text list "EncoderแกนX (เบิกจ่าย)": 0 '0'; 1 '5935'; 2 '9155'; 3 '12375'; 4 '15595'; 5 '18815'; 6 '22035'; 7 '25255'; 8 '28475'; 9 '31695'; 10 '34915'; 11 '38135'; 12 '41355'; 13 '44575'; 14 '52483'; 15 '55703'; 16 '58923'; 17 '62143'; 18 '65363'; 19 '68583'; 20 '71803'; 21 '75023'; 22 '78243'; 23 '81463'; 24 '84683'; 25 '87903'; 26 '91123'; 27 '5935'; 28 '9155'; 29 '12375'; 30 '15595'; 31 '18815'; 32 '22035'; 33 '25255'; 34 '28475'; 35 '31695'; 36 '34915'; 37 '38135'; 38 '41355'; 39 '44575'; 40 '52483'; 41 '55703'; 42 '58923'; 43 '62143'; 44 '65363'; 45 '68583'; 46 '71803'; 47 '75023'; 48 '78243'; 49 '81463'; 50 '84683'; 51 '87903'; 52 '91123'; 53 '5935'; 54 '9155'; 55 '12375'; 56 '15595'; 57 '18815'; 58 '22035'; 59 '25255'; 60 '28475'; 61 '31695'; 62 '34915'; 63 '38135'; 64 '41355'; 65 '44575'; 66 '52483'; 67 '55703'; 68 '58923'; 69 '62143'; 70 '65363'; 71 '68583'; 72 '71803'; 73 '75023'; 74 '78243'; 75 '81463'; 76 '84683'; 77 '87903'; 78 '91123'; 79 '5935'; 80 '9155'; 81 '12375'; 82 '15595'; 83 '18815'; 84 '22035'; 85 '25255'; 86 '28475'; 87 '31695'; 88 '34915'; 89 '38135'; 90 '41355'; 91 '44575'; 92 '52483'; 93 '55703'; 94 '58923'; 95 '62143'; 96 '65363'; 97 '68583'; 98 '71803'; 99 '75023'; 100 '78243'; 101 '81463'; 102 '84683'; 103 '87903'; 104 '91123'; 105 '5935'; 106 '9155'; 107 '12375'; 108 '15595'; 109 '18815'; 110 '22035'; 111 '25255'; 112 '28475'; 113 '31695'; 114 '34915'; 115 '38135'; 116 '41355'; 117 '44575'; 118 '52483'; 119 '55703'; 120 '58923'; 121 '62143'; 122 '65363'; 123 '68583'; 124 '71803'; 125 '75023'; 126 '78243'; 127 '81463'; 128 '84683'; 129 '87903'; 130 '91123'; 131 '5935'; 132 '9155'; 133 '12375'; 134 '15595'; 135 '18815'; 136 '22035'; 137 '25255'; 138 '28475'; 139 '31695'; 140 '34915'; 141 '38135'; 142 '41355'; 143 '44575'; 144 '52483'; 145 '55703'; 146 '58923'; 147 '62143'; 148 '65363'; 149 '68583'; 150 '71803'; 151 '75023'; 152 '78243'; 153 '81463'; 154 '84683'; 155 '87903'; 156 '91123'; 157 '5935'; 158 '9155'; 159 '12375'; 160 '15595'; 161 '18815'; 162 '22035'; 163 '25255'; 164 '28475'; 165 '31695'; 166 '34915'; 167 '38135'; 168 '41355'; 169 '44575'; 170 '52483'; 171 '55703'; 172 '58923'; 173 '62143'; 174 '65363'; 175 '68583'; 176 '71803'; 177 '75023'; 178 '78243'; 179 '81463'; 180 '84683'; 181 '87903'; 182 '91123'; 183 '5935'; 184 '9155'; 185 '12375'; 186 '15595'; 187 '18815'; 188 '22035'; 189 '25255'; 190 '28475'; 191 '31695'; 192 '34915'; 193 '38135'; 194 '41355'; 195 '44575'; 196 '52483'; 197 '55703'; 198 '58923'; 199 '62143'; 200 '65363'; 201 '68583'; 202 '71803'; 203 '75023'; 204 '78243'; 205 '81463'; 206 '84683'; 207 '87903'; 208 '91123'; 209 '5935'; 210 '9155'; 211 '12375'; 212 '15595'; 213 '18815'; 214 '22035'; 215 '25255'; 216 '28475'; 217 '31695'; 218 '34915'; 219 '38135'; 220 '41355'; 221 '44575'; 222 '52483'; 223 '55703'; 224 '58923'; 225 '62143'; 226 '65363'; 227 '68583'; 228 '71803'; 229 '75023'; 230 '78243'; 231 '81463'; 232 '84683'; 233 '87903'; 234 '91123'; 235 '5935'; 236 '9155'; 237 '12375'; 238 '15595'; 239 '18815'; 240 '22035'; 241 '25255'; 242 '28475'; 243 '31695'; 244 '34915'; 245 '38135'; 246 '41355'; 247 '44575'; 248 '52483'; 249 '55703'; 250 '58923'; 251 '62143'; 252 '65363'; 253 '68583'; 254 '71803'; 255 '75023'; 256 '78243'; 257 '81463'; 258 '84683'; 259 '87903'; 260 '91123'; 261 '5935'; 262 '9155'; 263 '12375'; 264 '15595'; 265 '18815'; 266 '22035'; 267 '25255'; 268 '28475'; 269 '31695'; 270 '34915'; 271 '38135'; 272 '41355'; 273 '44575'; 274 '52483'; 275 '55703'; 276 '58923'; 277 '62143'; 278 '65363'; 279 '68583'; 280 '71803'; 281 '75023'; 282 '78243'; 283 '81463'; 284 '84683'; 285 '87903'; 286 '91123'; 287 '5935'; 288 '9155'; 289 '12375'; 290 '15595'; 291 '18815'; 292 '22035'; 293 '25255'; 294 '28475'; 295 '31695'; 296 '34915'; 297 '38135'; 298 '41355'; 299 '44575'; 300 '52483'; 301 '55703'; 302 '58923'; 303 '62143'; 304 '65363'; 305 '68583'; 306 '71803'; 307 '75023'; 308 '78243'; 309 '81463'; 310 '84683'; 311 '87903'; 312 '91123'; 313 '5935'; 314 '9155'; 315 '12375'; 316 '15595'; 317 '18815'; 318 '22035'; 319 '25255'; 320 '28475'; 321 '31695'; 322 '34915'; 323 '38135'; 324 '41355'; 325 '44575'; 326 '52483'; 327 '55703'; 328 '58923'; 329 '62143'; 330 '65363'; 331 '68583'; 332 '71803'; 333 '75023'; 334 '78243'; 335 '81463'; 336 '84683'; 337 '87903'; 338 '91123'; 339 '5935'; 340 '9155'; 341 '12375'; 342 '15595'; 343 '18815'; 344 '22035'; 345 '25255'; 346 '28475'; 347 '31695'; 348 '34915'; 349 '38135'; 350 '41355'; 351 '44575'; 352 '52483'; 353 '55703'; 354 '58923'; 355 '62143'; 356 '65363'; 357 '68583'; 358 '71803'; 359 '75023'; 360 '78243'; 361 '81463'; 362 '84683'; 363 '87903'; 364 '91123'; 365 '5935'; 366 '9155'; 367 '12375'; 368 '15595'; 369 '18815'; 370 '22035'; 371 '25255'; 372 '28475'; 373 '31695'; 374 '34915'; 375 '38135'; 376 '41355'; 377 '44575'; 378 '52483'; 379 '55703'; 380 '58923'; 381 '62143'; 382 '65363'; 383 '68583'; 384 '71803'; 385 '75023'; 386 '78243'; 387 '81463'; 388 '84683'; 389 '87903'; 390 '91123'; 391 '5935'; 392 '9155'; 393 '12375'; 394 '15595'; 395 '18815'; 396 '22035'; 397 '25255'; 398 '28475'; 399 '31695'; 400 '34915'; 401 '38135'; 402 '41355'; 403 '44575'; 404 '52483'; 405 '55703'; 406 '58923'; 407 '62143'; 408 '65363'; 409 '68583'; 410 '71803'; 411 '75023'; 412 '78243'; 413 '81463'; 414 '84683'; 415 '87903'; 416 '91123'; 417 '5935'; 418 '9155'; 419 '12375'; 420 '15595'; 421 '18815'; 422 '22035'; 423 '25255'; 424 '28475'; 425 '31695'; 426 '34915'; 427 '38135'; 428 '41355'; 429 '44575'; 430 '52483'; 431 '55703'; 432 '58923'; 433 '62143'; 434 '65363'; 435 '68583'; 436 '71803'; 437 '75023'; 438 '78243'; 439 '81463'; 440 '84683'; 441 '87903'; 442 '91123'; 443 '5935'; 444 '9155'; 445 '12375'; 446 '15595'; 447 '18815'; 448 '22035'; 449 '25255'; 450 '28475'; 451 '31695'; 452 '34915'; 453 '38135'; 454 '41355'; 455 '44575'; 456 '52483'; 457 '55703'; 458 '58923'; 459 '62143'; 460 '65363'; 461 '68583'; 462 '71803'; 463 '75023'; 464 '78243'; 465 '81463'; 466 '84683'; 467 '87903'; 468 '91123'; 469 '5935'; 470 '9155'; 471 '12375'; 472 '15595'; 473 '18815'; 474 '22035'; 475 '25255'; 476 '28475'; 477 '31695'; 478 '34915'; 479 '38135'; 480 '41355'; 481 '44575'; 482 '52483'; 483 '55703'; 484 '58923'; 485 '62143'; 486 '65363'; 487 '68583'; 488 '71803'; 489 '75023'; 490 '78243'; 491 '81463'; 492 '84683'; 493 '87903'; 494 '91123'

text list "Textlist_ScreenName": 1 'PROCESS OVERVIEW'; 5 'ALARMS'; 20 'ORDER'; 10 'SETTING'

text list "จัดเก็บ Motor speed1,2": 0 '0'; 1 '500'

text list "จัดเก็บ Current 1,2": 0 '0'; 1 '6'

text list "จัดเก็บ Power 1,2": 0 '0'; 1 '270'

text list "จัดเก็บVoltage 1,2": 0 '0'; 1 '66'

text list "จัดเก็บ Motor speed3": 0 '0'; 2 '1500'

text list "จัดเก็บ Current 3": 0 '0'; 2 '6'

text list "จัดเก็บ Power 3": 0 '0'; 2 '270'

text list "จัดเก็บVoltage 3": 0 '0'; 2 '66'

text list "เบิกจ่าย Motor speed1,2": 0 '0'; 1 '500'

text list "เบิกจ่าย Current 1,2": 0 '0'; 1 '6'

text list "เบิกจ่าย Power 1,2": 0 '0'; 1 '270'

text list "เบิกจ่ายVoltage 1,2": 0 '0'; 1 '66'

text list "เบิกจ่าย Motor speed3": 0 '0'; 2 '1500'

text list "เบิกจ่าย Current 3": 0 '0'; 2 '6'

text list "เบิกจ่าย Power 3": 0 '0'; 2 '270'

text list "เบิกจ่ายVoltage 3": 0 '0'; 2 '66'

text list "Status1": 0 'Stop'; 1 'Running'

graphic list "GriphList_Button_Start": 0 '-play-button-off'; 1 '-button-96-on'

graphic list "GriphList_Button_Setting": 0 'setting-green-off'; 1 'settings-96-off'

graphic list "GriphList_Button_Alarms": 0 'arning-96-off'; 1 'warning-96-on'

graphic list "GriphList_Button_Order": 0 'order-off'; 1 'order'

graphic list "GriphList_Button_Overview": 0 'overview-off'; 1 'overview-on'

PopupScreen "Confirm" 500x250
   TextField "Template_Text field_1" at 72,8 size 209x37; Text 'ยืนยันการสั่งซื้อ'
   Button "Button_1" at 426,9 size 64x32; TextOff 'X'
      on Click: function_efd93a16("Confirm", 0, 0, 0, -1, 1)
   GraphicView "Template_Graphic view_1" at 8,8 size 45x40; Picture "bell"
   GraphicView "Template_Graphic view_2" at 152,66 size 187x166; Picture "accept"

PopupScreen "ช่องยานี้เต็มแล้ว" 500x250
   TextField "Template_Text field_1" at 72,8 size 22x37; Text 'Text'
   Button "Button_1" at 426,9 size 64x32; TextOff 'X'
      on Click: function_efd93a16("ช่องยานี้เต็มแล้ว", 0, 0, 0, -1, 1)
   GraphicView "Template_Graphic view_1" at 8,8 size 45x40; Picture "bell"
   GraphicView "Template_Graphic view_2" at 152,66 size 187x166; Picture "close"

PopupScreen "จัดเก็บยาเสร็จสิ้น" 500x250
   TextField "Template_Text field_1" at 72,8 size 227x37; Text 'จัดเก็บยาเสร็จสิ้น'
   Button "Button_1" at 426,9 size 64x32; TextOff 'X'
      on Click: function_efd93a16("จัดเก็บยาเสร็จสิ้น", 0, 0, 0, -1, 1)
   GraphicView "Template_Graphic view_1" at 8,8 size 45x40; Picture "bell"
   GraphicView "Template_Graphic view_2" at 152,66 size 187x166; Picture "accept"

Template "Template" 800x480
   TextField "Template_Text field_1" at 200,12 size 394x37; Text 'MAIN-PHARMACY SYSTEM'
   HTMLBrowser "Template_HTML browser_1" at 12,123 size 648x344
   DateTimeField "Template_Date/time field_1" at 320,43 size 131x26
   GraphicView "Template_Graphic view_7" at -1,0 size 110x139; Picture "MTET-Photoroom"
   GraphicView "Template_Graphic view_6" at 672,0 size 98x107; Picture "channels4_profile-Photoroom"
   TextField "Template_Text field_3" at 86,82 size 145x32; Text 'SYSTEM :'

Template "ORDER" 800x480
   TextField "Template_Text field_1" at 179,16 size 495x37; Text 'Medicine Retrieval System Screen'
   SymbolicIOField "Symbolic I/O field_1" at 376,204 size 386x72; TextOn '1'; TextOff '0'; TextList "SelectedMedicine"
      ProcessValue <- "แสดงชื่อยา"
      Appearance <- "แสดงชื่อยา"
   DateTimeField "Template_Date/time field_1" at 669,16 size 131x26
   Button "Button_2" at 368,77 size 400x56; TextOff 'Text'
   TextField "Template_Text field_2" at 367,88 size 401x32; Text 'ชื่อเวชภัณฑ์ (Medication Name):'
   Button "Button_1" at 368,137 size 400x56; TextOff 'Text'
   TextField "Template_Text field_3" at 382,148 size 214x32; Text 'รายการยาที่เลือก :'
   TextField "Template_Text field_4" at 616,147 size 20x32; Text 'Text'
   GraphicView "Template_Graphic view_1" at 21,68 size 72x64; Picture "Med"
   GraphicView "Template_Graphic view_2" at 25,134 size 65x58; Picture "tube"
   GraphicView "Template_Graphic view_3" at 25,202 size 63x56; Picture "vitamins"
   GraphicView "Template_Graphic view_4" at 23,269 size 64x57; Picture "medicine-pills"
   Button "Template_Button_3" at 368,368 size 192x88; TextOff 'CLEAR'
   GraphicView "Template_Graphic view_6" at 574,246 size 146x147; Picture "channels4_profile-Photoroom"
   GraphicView "Template_Graphic view_7" at 408,264 size 182x179; Picture "MTET-Photoroom"
   Button "Button_4" at 16,64 size 320x64; TextOff 'ยาแก้ปวด / ลดไข้'
      on Press: ActivateScreen("4_ORDER", 0)
   Button "Button_5" at 17,131 size 320x64; TextOff 'ยาทาภายนอก / ผิวหนัง'
      on Press: ActivateScreen("4_ORDER", 0)
   Button "Button_6" at 17,198 size 320x64; TextOff 'วิตามิน / อาหารเสริม'
      on Press: ActivateScreen("4_ORDER", 0)
   Button "Button_7" at 19,265 size 320x64; TextOff 'กลุ่มยาระบบทางเดินอาหาร'
      on Press: ActivateScreen("4_ORDER", 0)
   Button "Button_3" at 19,332 size 320x64; TextOff 'กลุ่มยาระบบทางเดินอาหาร'
      on Press: ActivateScreen("4_ORDER", 0)

Template "Template_2" 800x480
   TextField "Template_Text field_1" at 200,10 size 394x37; Text 'MAIN-PHARMACY SYSTEM'
   TextField "Template_Text field_2" at 81,80 size 145x32; Text 'SYSTEM :'
   DateTimeField "Template_Date/time field_1" at 328,44 size 131x26

Template "SETTING" 800x480
   DateTimeField "Template_Date/time field_1" at 98,37 size 131x26
   TextField "Template_Text field_2" at 448,312 size 20x32; Text 'Text'
   GraphicView "Template_Graphic view_7" at 21,5 size 87x90; Picture "channels4_profile-Photoroom"
   Button "Button_3" at 224,26 size 343x48; TextOff 'Text'
   TextField "Template_Text field_3" at 264,32 size 285x37; Text 'SYSTEM Animation'

Template "Alarms" 800x480
   DateTimeField "Template_Date/time field_1" at 648,32 size 131x26
   TextField "Template_Text field_2" at 448,312 size 20x32; Text 'Text'
   GraphicView "Template_Graphic view_7" at 21,5 size 87x90; Picture "channels4_profile-Photoroom"
   Button "Button_3" at 224,26 size 343x48; TextOff 'Text'
   TextField "Template_Text field_3" at 264,32 size 256x37; Text 'SYSTEM ALARMS'

Template "property HMI data" 800x480
   DateTimeField "Template_Date/time field_1" at 648,32 size 131x26
   GraphicView "Template_Graphic view_7" at 21,5 size 87x90; Picture "channels4_profile-Photoroom"
   Button "Button_3" at 224,26 size 343x48; TextOff 'Text'
   TextField "Template_Text field_1" at 254,31 size 273x37; Text 'property HMI data'
   TextField "Template_Text field_5" at 13,212 size 143x17; Text 'X AXIS ( Horizontall )'
   TextField "Template_Text field_6" at 27,227 size 57x17; Text 'Position'
   Button "Button_1" at 16,165 size 183x40; TextOff 'Text'
   TextField "Template_Text field_7" at 20,172 size 173x25; Text 'SERVO POSITION'
   TextField "Template_Text field_4" at 13,341 size 126x17; Text 'Y AXIS ( Verticall )'
   TextField "Template_Text field_8" at 27,356 size 57x17; Text 'Position'
   Button "Button_2" at 297,165 size 127x32; TextOff 'Text'
   TextField "Template_Text field_9" at 305,170 size 110x22; Text 'SERVO DATA'
   Button "Button_5" at 20,98 size 79x32; TextOff 'Text'
   TextField "Template_Text field_38" at 17,107 size 85x14; Text 'SEQUENCE STEP'
   TextField "Template_Text field_11" at 144,258 size 28x17; Text 'mm'
   TextField "Template_Text field_12" at 144,387 size 28x17; Text 'mm'
   Button "Button_4" at 408,87 size 183x64; TextOff 'Text'

Template "Status system" 800x480
   TextField "Template_Text field_1" at 256,8 size 318x37; Text 'Status System Screen'
   Button "Template_Button_1" at 16,80 size 184x48; TextOff 'เบิกจ่าย ( Retrieval )'
   Button "Template_Button_2" at 220,79 size 184x48; TextOff 'จัดเก็บ ( Storage )'
   Circle "Template_Circle_1" at 16,450 size 24x24
      Appearance <- "Output Status2"
   Circle "Template_Circle_2" at 218,450 size 24x24
      Appearance <- "Output Status1"
   SymbolicIOField "Template_Symbolic I/O field_1" at 323,450 size 82x23; TextOn '1'; TextOff '0'; TextList "Status1"
      ProcessValue <- "Output Status1"
   SymbolicIOField "Template_Symbolic I/O field_2" at 120,450 size 82x23; TextOn '1'; TextOff '0'; TextList "Status1"
      ProcessValue <- "Output Status2"
   HTMLBrowser "Template_HTML browser_1" at 424,159 size 352x248
      Address <- "Video_URL"
   TextField "Template_Text field_4" at 616,147 size 20x32; Text 'Text'
   TextField "Template_Text field_3" at 464,88 size 322x22; Text 'คลิปการทำงาน : การเบิกจ่าย / การจัดเก็บ'
   DateTimeField "Template_Date/time field_1" at 642,16 size 131x26
   GraphicView "Template_Graphic view_6" at 95,-2 size 73x67; Picture "channels4_profile-Photoroom"
   GraphicView "Template_Graphic view_7" at 2,2 size 102x106; Picture "MTET-Photoroom"
   TextField "Template_Text field_2" at 32,455 size 96x14; Text 'MACHINE STATUS :'
   TextField "Template_Text field_5" at 235,455 size 96x14; Text 'MACHINE STATUS :'
   GraphicView "Template_Graphic view_1" at 432,78 size 47x43; Picture "video-clip"
   GraphicView "Template_Graphic view_2" at 229,81 size 47x43; Picture "storage-room"
   GraphicView "Template_Graphic view_3" at 23,82 size 47x43; Picture "shopping-cart"

Template "Keep_1" 800x480
   TextField "Template_Text field_1" at 200,10 size 394x37; Text 'MAIN-PHARMACY SYSTEM'
   TextField "Template_Text field_2" at 122,88 size 384x37; Text 'Pharmacy Storage System'
   DateTimeField "Template_Date/time field_1" at 328,44 size 131x26

screen "LOGIN" 800x480, template "Template"
   Button "Button_2" at 668,96 size 128x72; TextOff 'LOGIN'; Authorization "Admin"
      on Activate: function_a2a04561(); ActivateScreen("1_OVERVIEW_1", 0)
   Button "Button_6" at 668,398 size 128x72; TextOn 'LOGOUT'; TextOff 'LOGOUT'
      on Activate: function_f23ef4c9(); ActivateScreen("LOGIN", 0)
   GraphicView "Template_Graphic view_1" at 672,107 size 54x48; Picture "NEW_HOME"
   GraphicView "Template_Graphic view_5" at 672,413 size 54x48; Picture "logout"

screen "1_2" 800x480, template "Template_2"
   Button "Button_1" at 40,240 size 120x40; TextOff 'Oxytocin'
      on Click: ActivateScreen("4_ORDER", 0); SetTag("Selected_URL", 'file:///C:/ASRS_Video/clip341.html')
      on Activate: SetTag("Selected_Medicine", 341)
      on Release: SetTag("ยา 341", 0)
      on Press: SetTag("ยา 341", 1)
   Button "Button_10" at 38,415 size 120x40; TextOff 'Nifedipine'
      on Click: ActivateScreen("4_ORDER", 0); SetTag("Selected_URL", 'file:///C:/ASRS_Video/clip346.html')
      on Activate: SetTag("Selected_Medicine", 346)
      on Release: SetTag("ยา 346", 0)
      on Press: SetTag("ยา 346", 1)
   Button "Button_2" at 189,240 size 120x40; TextOff 'Misoprostol'
      on Click: ActivateScreen("4_ORDER", 0); SetTag("Selected_URL", 'file:///C:/ASRS_Video/clip342.html')
      on Activate: SetTag("Selected_Medicine", 342)
      on Release: SetTag("ยา 342", 0)
      on Press: SetTag("ยา 342", 1)
   Button "Button_3" at 190,415 size 120x40; TextOff 'Terbutaline'
      on Click: ActivateScreen("4_ORDER", 0); SetTag("Selected_URL", 'file:///C:/ASRS_Video/clip347.html')
      on Activate: SetTag("Selected_Medicine", 347)
      on Release: SetTag("ยา 347", 0)
      on Press: SetTag("ยา 347", 1)
   Button "Button_4" at 340,240 size 120x40; TextOff 'Dinoprostone'
      on Click: ActivateScreen("4_ORDER", 0); SetTag("Selected_URL", 'file:///C:/ASRS_Video/clip343.html')
      on Activate: SetTag("Selected_Medicine", 343)
      on Release: SetTag("ยา 343", 0)
      on Press: SetTag("ยา 343", 1)
   Button "Button_5" at 340,416 size 120x40; TextOff 'Ferrous fumarate'
      on Click: ActivateScreen("4_ORDER", 0); SetTag("Selected_URL", 'file:///C:/ASRS_Video/clip348.html')
      on Activate: SetTag("Selected_Medicine", 348)
      on Release: SetTag("ยา 348", 0)
      on Press: SetTag("ยา 348", 1)
   Button "Button_6" at 492,416 size 120x40; TextOff 'Folic acid'
      on Click: ActivateScreen("4_ORDER", 0); SetTag("Selected_URL", 'file:///C:/ASRS_Video/clip349.html')
      on Activate: SetTag("Selected_Medicine", 349)
      on Release: SetTag("ยา 349", 0)
      on Press: SetTag("ยา 349", 1)
   Button "Button_7" at 492,240 size 120x40; TextOff 'Methylergometrine'
      on Click: ActivateScreen("4_ORDER", 0); SetTag("Selected_URL", 'file:///C:/ASRS_Video/clip344.html')
      on Activate: SetTag("Selected_Medicine", 344)
      on Release: SetTag("ยา 344", 0)
      on Press: SetTag("ยา 344", 1)
   Button "Button_8" at 644,240 size 120x40; TextOff 'Magnesium sulfate'
      on Click: ActivateScreen("4_ORDER", 0); SetTag("Selected_URL", 'file:///C:/ASRS_Video/clip345.html')
      on Activate: SetTag("Selected_Medicine", 345)
      on Release: SetTag("ยา 345", 0)
      on Press: SetTag("ยา 345", 1)
   Button "Button_11" at 645,416 size 120x40; TextOff 'Calcium carbonate'
      on Click: ActivateScreen("4_ORDER", 0); SetTag("Selected_URL", 'file:///C:/ASRS_Video/clip350.html')
      on Activate: SetTag("Selected_Medicine", 350)
      on Release: SetTag("ยา 350", 0)
      on Press: SetTag("ยา 350", 1)
   Button "Button_12" at 688,16 size 96x40; TextOff 'Next'
      on Press: ActivateScreen("2_2", 0)
   Button "Button_9" at 24,16 size 94x40; TextOff 'Back'
      on Press: ActivateScreen("4_ORDER", 0)
   GraphicView "Template_Graphic view_2" at 693,20 size 36x32; Picture "play"
   GraphicView "Template_Graphic view_1" at 27,19 size 36x32; Picture "fast-backward"
   GraphicView "Template_Graphic view_3" at 37,128 size 120x104; Picture "1_1"
   GraphicView "Template_Graphic view_4" at 191,129 size 120x104; Picture "2_1"
   GraphicView "Template_Graphic view_5" at 339,129 size 120x104; Picture "3_1"
   GraphicView "Template_Graphic view_6" at 493,129 size 120x104; Picture "4_1"
   GraphicView "Template_Graphic view_7" at 645,129 size 120x104; Picture "5_1"
   GraphicView "Template_Graphic view_8" at 38,305 size 120x104; Picture "6_1"
   GraphicView "Template_Graphic view_9" at 189,304 size 120x112; Picture "7_1"
   GraphicView "Template_Graphic view_10" at 351,307 size 96x104; Picture "8_1"
   GraphicView "Template_Graphic view_11" at 497,304 size 120x112; Picture "9_1"
   GraphicView "Template_Graphic view_12" at 645,304 size 120x104; Picture "10_1"
   TextField "Template_Text field_2" at 201,80 size 20x32; Text '1'

screen "2_2" 800x480, template "Template_2"
   Button "Button_1" at 38,239 size 120x40; TextOff 'Ethinylestradiol'
      on Click: ActivateScreen("4_ORDER", 0); SetTag("Selected_URL", 'file:///C:/ASRS_Video/clip351.html')
      on Activate: SetTag("Selected_Medicine", 351)
      on Release: SetTag("ยา 351", 0)
      on Press: SetTag("ยา 351", 1)
   Button "Button_9" at 688,16 size 96x40; TextOff 'Next'
      on Press: ActivateScreen("3_2", 0)
   Button "Button_10" at 38,415 size 120x40; TextOff 'Letrozole'
      on Click: ActivateScreen("4_ORDER", 0); SetTag("Selected_URL", 'file:///C:/ASRS_Video/clip356.html')
      on Activate: SetTag("Selected_Medicine", 356)
      on Release: SetTag("ยา 356", 0)
      on Press: SetTag("ยา 356", 1)
   Button "Button_2" at 189,240 size 120x40; TextOff 'Levonorgestrel'
      on Click: ActivateScreen("4_ORDER", 0); SetTag("Selected_URL", 'file:///C:/ASRS_Video/clip352.html')
      on Activate: SetTag("Selected_Medicine", 352)
      on Release: SetTag("ยา 352", 0)
      on Press: SetTag("ยา 352", 1)
   Button "Button_3" at 190,415 size 120x40; TextOff 'Tamoxifen'
      on Click: ActivateScreen("4_ORDER", 0); SetTag("Selected_URL", 'file:///C:/ASRS_Video/clip357.html')
      on Activate: SetTag("Selected_Medicine", 357)
      on Release: SetTag("ยา 357", 0)
      on Press: SetTag("ยา 357", 1)
   Button "Button_4" at 340,240 size 120x40; TextOff 'Medroxyprogesterone'
      on Click: ActivateScreen("4_ORDER", 0); SetTag("Selected_URL", 'file:///C:/ASRS_Video/clip353.html')
      on Activate: SetTag("Selected_Medicine", 353)
      on Release: SetTag("ยา 353", 0)
      on Press: SetTag("ยา 353", 1)
   Button "Button_5" at 340,416 size 120x40; TextOff 'Anastrozole'
      on Click: ActivateScreen("4_ORDER", 0); SetTag("Selected_URL", 'file:///C:/ASRS_Video/clip358.html')
      on Activate: SetTag("Selected_Medicine", 358)
      on Release: SetTag("ยา 358", 0)
      on Press: SetTag("ยา 358", 1)
   Button "Button_6" at 492,416 size 120x40; TextOff 'Exemestane'
      on Click: ActivateScreen("4_ORDER", 0); SetTag("Selected_URL", 'file:///C:/ASRS_Video/clip359.html')
      on Activate: SetTag("Selected_Medicine", 359)
      on Release: SetTag("ยา 359", 0)
      on Press: SetTag("ยา 359", 1)
   Button "Button_7" at 492,240 size 120x40; TextOff 'Norethisterone'
      on Click: ActivateScreen("4_ORDER", 0); SetTag("Selected_URL", 'file:///C:/ASRS_Video/clip354.html')
      on Activate: SetTag("Selected_Medicine", 354)
      on Release: SetTag("ยา 354", 0)
      on Press: SetTag("ยา 354", 1)
   Button "Button_8" at 644,240 size 120x40; TextOff 'Clomiphene citrate'
      on Click: ActivateScreen("4_ORDER", 0); SetTag("Selected_URL", 'file:///C:/ASRS_Video/clip355.html')
      on Activate: SetTag("Selected_Medicine", 355)
      on Release: SetTag("ยา 355", 0)
      on Press: SetTag("ยา 355", 1)
   Button "Button_11" at 645,416 size 120x40; TextOff 'Leuprolide'
      on Click: ActivateScreen("4_ORDER", 0); SetTag("Selected_URL", 'file:///C:/ASRS_Video/clip360.html')
      on Activate: SetTag("Selected_Medicine", 360)
      on Release: SetTag("ยา 360", 0)
      on Press: SetTag("ยา 360", 1)
   Button "Button_12" at 24,16 size 94x40; TextOff 'Back'
      on Press: ActivateScreen("1_2", 0)
   GraphicView "Template_Graphic view_1" at 693,20 size 36x32; Picture "play"
   GraphicView "Template_Graphic view_2" at 27,19 size 36x32; Picture "fast-backward"
   GraphicView "Template_Graphic view_3" at 37,128 size 120x104; Picture "11_1"
   GraphicView "Template_Graphic view_4" at 191,129 size 120x104; Picture "12_1"
   GraphicView "Template_Graphic view_5" at 339,129 size 120x104; Picture "13_1"
   GraphicView "Template_Graphic view_6" at 493,129 size 120x104; Picture "14_1"
   GraphicView "Template_Graphic view_7" at 645,129 size 120x104; Picture "15_1"
   GraphicView "Template_Graphic view_8" at 38,305 size 120x104; Picture "16_1"
   GraphicView "Template_Graphic view_9" at 189,304 size 120x112; Picture "17_1"
   GraphicView "Template_Graphic view_10" at 351,307 size 96x104; Picture "118"
   GraphicView "Template_Graphic view_11" at 497,304 size 120x112; Picture "19_1"
   GraphicView "Template_Graphic view_12" at 645,304 size 120x104; Picture "20_1"
   TextField "Template_Text field_2" at 201,80 size 20x32; Text '2'

screen "3_2" 800x480, template "Template_2"
   Button "Button_1" at 38,239 size 120x40; TextOff 'Goserelin'
      on Click: ActivateScreen("4_ORDER", 0); SetTag("Selected_URL", 'file:///C:/ASRS_Video/clip361.html')
      on Activate: SetTag("Selected_Medicine", 361)
      on Release: SetTag("ยา 361", 0)
      on Press: SetTag("ยา 361", 1)
   Button "Button_9" at 688,16 size 96x40; TextOff 'Next'
      on Press: ActivateScreen("4_2", 0)
   Button "Button_10" at 38,415 size 120x40; TextOff 'Oxybutynin'
      on Click: ActivateScreen("4_ORDER", 0); SetTag("Selected_URL", 'file:///C:/ASRS_Video/clip366.html')
      on Activate: SetTag("Selected_Medicine", 366)
      on Release: SetTag("ยา 366", 0)
      on Press: SetTag("ยา 366", 1)
   Button "Button_2" at 189,240 size 120x40; TextOff 'Finasteride'
      on Click: ActivateScreen("4_ORDER", 0); SetTag("Selected_URL", 'file:///C:/ASRS_Video/clip362.html')
      on Activate: SetTag("Selected_Medicine", 362)
      on Release: SetTag("ยา 362", 0)
      on Press: SetTag("ยา 362", 1)
   Button "Button_3" at 190,415 size 120x40; TextOff 'Tolterodine'
      on Click: ActivateScreen("4_ORDER", 0); SetTag("Selected_URL", 'file:///C:/ASRS_Video/clip367.html')
      on Activate: SetTag("Selected_Medicine", 367)
      on Release: SetTag("ยา 367", 0)
      on Press: SetTag("ยา 367", 1)
   Button "Button_4" at 340,240 size 120x40; TextOff 'Dutasteride'
      on Click: ActivateScreen("4_ORDER", 0); SetTag("Selected_URL", 'file:///C:/ASRS_Video/clip363.html')
      on Activate: SetTag("Selected_Medicine", 363)
      on Release: SetTag("ยา 363", 0)
      on Press: SetTag("ยา 363", 1)
   Button "Button_5" at 340,416 size 120x40; TextOff 'Solifenacin'
      on Click: ActivateScreen("4_ORDER", 0); SetTag("Selected_URL", 'file:///C:/ASRS_Video/clip368.html')
      on Activate: SetTag("Selected_Medicine", 368)
      on Release: SetTag("ยา 368", 0)
      on Press: SetTag("ยา 368", 1)
   Button "Button_6" at 492,416 size 120x40; TextOff 'Mirabegron'
      on Click: ActivateScreen("4_ORDER", 0); SetTag("Selected_URL", 'file:///C:/ASRS_Video/clip369.html')
      on Activate: SetTag("Selected_Medicine", 369)
      on Release: SetTag("ยา 369", 0)
      on Press: SetTag("ยา 369", 1)
   Button "Button_7" at 492,240 size 120x40; TextOff 'Tamsulosin'
      on Click: ActivateScreen("4_ORDER", 0); SetTag("Selected_URL", 'file:///C:/ASRS_Video/clip364.html')
      on Activate: SetTag("Selected_Medicine", 364)
      on Release: SetTag("ยา 364", 0)
      on Press: SetTag("ยา 364", 1)
   Button "Button_8" at 644,240 size 120x40; TextOff 'Alfuzosin'
      on Click: ActivateScreen("4_ORDER", 0); SetTag("Selected_URL", 'file:///C:/ASRS_Video/clip365.html')
      on Activate: SetTag("Selected_Medicine", 365)
      on Release: SetTag("ยา 365", 0)
      on Press: SetTag("ยา 365", 1)
   Button "Button_11" at 645,416 size 120x40; TextOff 'Potassium citrate'
      on Click: ActivateScreen("4_ORDER", 0); SetTag("Selected_URL", 'file:///C:/ASRS_Video/clip370.html')
      on Activate: SetTag("Selected_Medicine", 370)
      on Release: SetTag("ยา 370", 0)
      on Press: SetTag("ยา 370", 1)
   Button "Button_12" at 24,16 size 94x40; TextOff 'Back'
      on Press: ActivateScreen("2_2", 0)
   GraphicView "Template_Graphic view_1" at 693,20 size 36x32; Picture "play"
   GraphicView "Template_Graphic view_2" at 27,19 size 36x32; Picture "fast-backward"
   GraphicView "Template_Graphic view_3" at 37,128 size 120x104; Picture "21_1"
   GraphicView "Template_Graphic view_4" at 191,129 size 120x104; Picture "22_1"
   GraphicView "Template_Graphic view_5" at 339,129 size 120x104; Picture "23_1"
   GraphicView "Template_Graphic view_6" at 493,129 size 120x104; Picture "24_1"
   GraphicView "Template_Graphic view_7" at 645,129 size 120x104; Picture "25_1"
   GraphicView "Template_Graphic view_8" at 38,305 size 120x104; Picture "26_1"
   GraphicView "Template_Graphic view_9" at 189,304 size 120x112; Picture "27_1"
   GraphicView "Template_Graphic view_10" at 351,307 size 96x104; Picture "28_1"
   GraphicView "Template_Graphic view_11" at 497,304 size 120x112; Picture "29_1"
   GraphicView "Template_Graphic view_12" at 645,304 size 120x104; Picture "30_1"
   TextField "Template_Text field_2" at 201,80 size 20x32; Text '3'

screen "4_2" 800x480, template "Template_2"
   Button "Button_1" at 38,239 size 120x40; TextOff 'Sodium bicarbonate'
      on Click: ActivateScreen("4_ORDER", 0); SetTag("Selected_URL", 'file:///C:/ASRS_Video/clip371.html')
      on Activate: SetTag("Selected_Medicine", 371)
      on Release: SetTag("ยา 371", 0)
      on Press: SetTag("ยา 371", 1)
   Button "Button_9" at 688,16 size 96x40; TextOff 'Next'
      on Press: ActivateScreen("5_2", 0)
   Button "Button_10" at 38,415 size 120x40; TextOff 'Ifosfamide'
      on Click: ActivateScreen("4_ORDER", 0); SetTag("Selected_URL", 'file:///C:/ASRS_Video/clip376.html')
      on Activate: SetTag("Selected_Medicine", 376)
      on Release: SetTag("ยา 376", 0)
      on Press: SetTag("ยา 376", 1)
   Button "Button_2" at 189,240 size 120x40; TextOff 'Nitrofurantoin'
      on Click: ActivateScreen("4_ORDER", 0); SetTag("Selected_URL", 'file:///C:/ASRS_Video/clip372.html')
      on Activate: SetTag("Selected_Medicine", 372)
      on Release: SetTag("ยา 372", 0)
      on Press: SetTag("ยา 372", 1)
   Button "Button_3" at 190,415 size 120x40; TextOff 'Chlorambucil'
      on Click: ActivateScreen("4_ORDER", 0); SetTag("Selected_URL", 'file:///C:/ASRS_Video/clip377.html')
      on Activate: SetTag("Selected_Medicine", 377)
      on Release: SetTag("ยา 377", 0)
      on Press: SetTag("ยา 377", 1)
   Button "Button_4" at 340,240 size 120x40; TextOff 'Fosfomycin'
      on Click: ActivateScreen("4_ORDER", 0); SetTag("Selected_URL", 'file:///C:/ASRS_Video/clip373.html')
      on Activate: SetTag("Selected_Medicine", 373)
      on Release: SetTag("ยา 373", 0)
      on Press: SetTag("ยา 373", 1)
   Button "Button_5" at 340,416 size 120x40; TextOff 'Melphalan'
      on Click: ActivateScreen("4_ORDER", 0); SetTag("Selected_URL", 'file:///C:/ASRS_Video/clip378.html')
      on Activate: SetTag("Selected_Medicine", 378)
      on Release: SetTag("ยา 378", 0)
      on Press: SetTag("ยา 378", 1)
   Button "Button_6" at 492,416 size 120x40; TextOff 'Busulfan'
      on Click: ActivateScreen("4_ORDER", 0); SetTag("Selected_URL", 'file:///C:/ASRS_Video/clip379.html')
      on Activate: SetTag("Selected_Medicine", 379)
      on Release: SetTag("ยา 379", 0)
      on Press: SetTag("ยา 379", 1)
   Button "Button_7" at 492,240 size 120x40; TextOff 'Methotrexate'
      on Click: ActivateScreen("4_ORDER", 0); SetTag("Selected_URL", 'file:///C:/ASRS_Video/clip374.html')
      on Activate: SetTag("Selected_Medicine", 374)
      on Release: SetTag("ยา 374", 0)
      on Press: SetTag("ยา 374", 1)
   Button "Button_8" at 644,240 size 120x40; TextOff 'Cyclophosphamide'
      on Click: ActivateScreen("4_ORDER", 0); SetTag("Selected_URL", 'file:///C:/ASRS_Video/clip375.html')
      on Activate: SetTag("Selected_Medicine", 375)
      on Release: SetTag("ยา 375", 0)
      on Press: SetTag("ยา 375", 1)
   Button "Button_11" at 645,416 size 120x40; TextOff 'Cytarabine'
      on Click: ActivateScreen("4_ORDER", 0); SetTag("Selected_URL", 'file:///C:/ASRS_Video/clip380.html')
      on Activate: SetTag("Selected_Medicine", 380)
      on Release: SetTag("ยา 380", 0)
      on Press: SetTag("ยา 380", 1)
   Button "Button_12" at 24,16 size 94x40; TextOff 'Back'
      on Press: ActivateScreen("3_2", 0)
   GraphicView "Template_Graphic view_1" at 693,20 size 36x32; Picture "play"
   GraphicView "Template_Graphic view_2" at 27,19 size 36x32; Picture "fast-backward"
   GraphicView "Template_Graphic view_3" at 37,128 size 120x104; Picture "31_1"
   GraphicView "Template_Graphic view_4" at 191,129 size 120x104; Picture "32_1"
   GraphicView "Template_Graphic view_5" at 339,129 size 120x104; Picture "33_1"
   GraphicView "Template_Graphic view_6" at 493,129 size 120x104; Picture "34_1"
   GraphicView "Template_Graphic view_7" at 645,129 size 120x104; Picture "35_1"
   GraphicView "Template_Graphic view_8" at 38,305 size 120x104; Picture "36_1"
   GraphicView "Template_Graphic view_9" at 189,304 size 120x112; Picture "37_1"
   GraphicView "Template_Graphic view_10" at 351,307 size 96x104; Picture "38_1"
   GraphicView "Template_Graphic view_11" at 497,304 size 120x112; Picture "39_1"
   GraphicView "Template_Graphic view_12" at 645,304 size 120x104; Picture "40_1"
   TextField "Template_Text field_2" at 201,80 size 20x32; Text '4'

screen "5_2" 800x480, template "Template_2"
   Button "Button_1" at 38,239 size 120x40; TextOff 'Fluorouracil'
      on Click: ActivateScreen("4_ORDER", 0); SetTag("Selected_URL", 'file:///C:/ASRS_Video/clip381.html')
      on Activate: SetTag("Selected_Medicine", 381)
      on Release: SetTag("ยา 381", 0)
      on Press: SetTag("ยา 381", 1)
   Button "Button_9" at 688,16 size 96x40; TextOff 'Next'
      on Press: ActivateScreen("6_2", 0)
   Button "Button_10" at 38,415 size 120x40; TextOff 'Epirubicin'
      on Click: ActivateScreen("4_ORDER", 0); SetTag("Selected_URL", 'file:///C:/ASRS_Video/clip386.html')
      on Activate: SetTag("Selected_Medicine", 386)
      on Release: SetTag("ยา 386", 0)
      on Press: SetTag("ยา 386", 1)
   Button "Button_2" at 189,240 size 120x40; TextOff 'Capecitabine'
      on Click: ActivateScreen("4_ORDER", 0); SetTag("Selected_URL", 'file:///C:/ASRS_Video/clip382.html')
      on Activate: SetTag("Selected_Medicine", 382)
      on Release: SetTag("ยา 382", 0)
      on Press: SetTag("ยา 382", 1)
   Button "Button_3" at 190,415 size 120x40; TextOff 'Bleomycin'
      on Click: ActivateScreen("4_ORDER", 0); SetTag("Selected_URL", 'file:///C:/ASRS_Video/clip387.html')
      on Activate: SetTag("Selected_Medicine", 387)
      on Release: SetTag("ยา 387", 0)
      on Press: SetTag("ยา 387", 1)
   Button "Button_4" at 340,240 size 120x40; TextOff 'Gemcitabine'
      on Click: ActivateScreen("4_ORDER", 0); SetTag("Selected_URL", 'file:///C:/ASRS_Video/clip383.html')
      on Activate: SetTag("Selected_Medicine", 383)
      on Release: SetTag("ยา 383", 0)
      on Press: SetTag("ยา 383", 1)
   Button "Button_5" at 340,416 size 120x40; TextOff 'Vincristine'
      on Click: ActivateScreen("4_ORDER", 0); SetTag("Selected_URL", 'file:///C:/ASRS_Video/clip388.html')
      on Activate: SetTag("Selected_Medicine", 388)
      on Release: SetTag("ยา 388", 0)
      on Press: SetTag("ยา 388", 1)
   Button "Button_6" at 492,416 size 120x40; TextOff 'Vinblastine'
      on Click: ActivateScreen("4_ORDER", 0); SetTag("Selected_URL", 'file:///C:/ASRS_Video/clip389.html')
      on Activate: SetTag("Selected_Medicine", 389)
      on Release: SetTag("ยา 389", 0)
      on Press: SetTag("ยา 389", 1)
   Button "Button_7" at 492,240 size 120x40; TextOff 'Doxorubicin'
      on Click: ActivateScreen("4_ORDER", 0); SetTag("Selected_URL", 'file:///C:/ASRS_Video/clip384.html')
      on Activate: SetTag("Selected_Medicine", 384)
      on Release: SetTag("ยา 384", 0)
      on Press: SetTag("ยา 384", 1)
   Button "Button_8" at 644,240 size 120x40; TextOff 'Daunorubicin'
      on Click: ActivateScreen("4_ORDER", 0); SetTag("Selected_URL", 'file:///C:/ASRS_Video/clip385.html')
      on Activate: SetTag("Selected_Medicine", 385)
      on Release: SetTag("ยา 385", 0)
      on Press: SetTag("ยา 385", 1)
   Button "Button_11" at 645,416 size 120x40; TextOff 'Paclitaxel'
      on Click: ActivateScreen("4_ORDER", 0); SetTag("Selected_URL", 'file:///C:/ASRS_Video/clip390.html')
      on Activate: SetTag("Selected_Medicine", 390)
      on Release: SetTag("ยา 390", 0)
      on Press: SetTag("ยา 390", 1)
   Button "Button_12" at 24,16 size 94x40; TextOff 'Back'
      on Press: ActivateScreen("4_2", 0)
   GraphicView "Template_Graphic view_1" at 693,20 size 36x32; Picture "play"
   GraphicView "Template_Graphic view_2" at 27,19 size 36x32; Picture "fast-backward"
   GraphicView "Template_Graphic view_3" at 37,128 size 120x104; Picture "41_1"
   GraphicView "Template_Graphic view_4" at 191,129 size 120x104; Picture "42_1"
   GraphicView "Template_Graphic view_5" at 339,129 size 120x104; Picture "43_1"
   GraphicView "Template_Graphic view_6" at 493,129 size 120x104; Picture "44_1"
   GraphicView "Template_Graphic view_7" at 645,129 size 120x104; Picture "45_1"
   GraphicView "Template_Graphic view_8" at 38,305 size 120x104; Picture "46_1"
   GraphicView "Template_Graphic view_9" at 189,304 size 120x112; Picture "47_1"
   GraphicView "Template_Graphic view_10" at 351,307 size 96x104; Picture "48_1"
   GraphicView "Template_Graphic view_11" at 497,304 size 120x112; Picture "49_1"
   GraphicView "Template_Graphic view_12" at 645,304 size 120x104; Picture "50_1"
   TextField "Template_Text field_2" at 201,80 size 20x32; Text '5'

screen "6_2" 800x480, template "Template_2"
   Button "Button_1" at 38,239 size 120x40; TextOff 'Docetaxel'
      on Click: ActivateScreen("4_ORDER", 0); SetTag("Selected_URL", 'file:///C:/ASRS_Video/clip391.html')
      on Activate: SetTag("Selected_Medicine", 391)
      on Release: SetTag("ยา 391", 0)
      on Press: SetTag("ยา 391", 1)
   Button "Button_9" at 688,16 size 96x40; TextOff 'Next'
      on Press: ActivateScreen("7_2", 0)
   Button "Button_10" at 38,415 size 120x40; TextOff 'Etoposide'
      on Click: ActivateScreen("4_ORDER", 0); SetTag("Selected_URL", 'file:///C:/ASRS_Video/clip396.html')
      on Activate: SetTag("Selected_Medicine", 396)
      on Release: SetTag("ยา 396", 0)
      on Press: SetTag("ยา 396", 1)
   Button "Button_2" at 188,238 size 120x40; TextOff 'Cisplatin'
      on Click: ActivateScreen("4_ORDER", 0); SetTag("Selected_URL", 'file:///C:/ASRS_Video/clip392.html')
      on Activate: SetTag("Selected_Medicine", 392)
      on Release: SetTag("ยา 392", 0)
      on Press: SetTag("ยา 392", 1)
   Button "Button_3" at 190,415 size 120x40; TextOff 'Topotecan'
      on Click: ActivateScreen("4_ORDER", 0); SetTag("Selected_URL", 'file:///C:/ASRS_Video/clip397.html')
      on Activate: SetTag("Selected_Medicine", 397)
      on Release: SetTag("ยา 397", 0)
      on Press: SetTag("ยา 397", 1)
   Button "Button_4" at 340,240 size 120x40; TextOff 'Carboplatin'
      on Click: ActivateScreen("4_ORDER", 0); SetTag("Selected_URL", 'file:///C:/ASRS_Video/clip393.html')
      on Activate: SetTag("Selected_Medicine", 393)
      on Release: SetTag("ยา 393", 0)
      on Press: SetTag("ยา 393", 1)
   Button "Button_5" at 340,416 size 120x40; TextOff 'Hydroxyurea'
      on Click: ActivateScreen("4_ORDER", 0); SetTag("Selected_URL", 'file:///C:/ASRS_Video/clip398.html')
      on Activate: SetTag("Selected_Medicine", 398)
      on Release: SetTag("ยา 398", 0)
      on Press: SetTag("ยา 398", 1)
   Button "Button_6" at 492,416 size 120x40; TextOff 'Mercaptopurine'
      on Click: ActivateScreen("4_ORDER", 0); SetTag("Selected_URL", 'file:///C:/ASRS_Video/clip399.html')
      on Activate: SetTag("Selected_Medicine", 399)
      on Release: SetTag("ยา 399", 0)
      on Press: SetTag("ยา 399", 1)
   Button "Button_7" at 492,240 size 120x40; TextOff 'Oxaliplatin'
      on Click: ActivateScreen("4_ORDER", 0); SetTag("Selected_URL", 'file:///C:/ASRS_Video/clip394.html')
      on Activate: SetTag("Selected_Medicine", 394)
      on Release: SetTag("ยา 394", 0)
      on Press: SetTag("ยา 394", 1)
   Button "Button_8" at 644,240 size 120x40; TextOff 'Irinotecan'
      on Click: ActivateScreen("4_ORDER", 0); SetTag("Selected_URL", 'file:///C:/ASRS_Video/clip395.html')
      on Activate: SetTag("Selected_Medicine", 395)
      on Release: SetTag("ยา 395", 0)
      on Press: SetTag("ยา 395", 1)
   Button "Button_11" at 645,416 size 120x40; TextOff 'Thioguanine'
      on Click: ActivateScreen("4_ORDER", 0); SetTag("Selected_URL", 'file:///C:/ASRS_Video/clip400.html')
      on Activate: SetTag("Selected_Medicine", 400)
      on Release: SetTag("ยา 400", 0)
      on Press: SetTag("ยา 400", 1)
   Button "Button_12" at 24,16 size 94x40; TextOff 'Back'
      on Press: ActivateScreen("5_2", 0)
   GraphicView "Template_Graphic view_1" at 693,20 size 36x32; Picture "play"
   GraphicView "Template_Graphic view_2" at 27,19 size 36x32; Picture "fast-backward"
   GraphicView "Template_Graphic view_3" at 37,128 size 120x104; Picture "51_1"
   GraphicView "Template_Graphic view_4" at 191,129 size 120x104; Picture "52_1"
   GraphicView "Template_Graphic view_5" at 339,129 size 120x104; Picture "53_1"
   GraphicView "Template_Graphic view_6" at 493,129 size 120x104; Picture "54_1"
   GraphicView "Template_Graphic view_7" at 645,129 size 120x104; Picture "55_1"
   GraphicView "Template_Graphic view_8" at 38,305 size 120x104; Picture "56_1"
   GraphicView "Template_Graphic view_9" at 189,304 size 120x112; Picture "57_1"
   GraphicView "Template_Graphic view_10" at 351,307 size 96x104; Picture "58_1"
   GraphicView "Template_Graphic view_11" at 497,304 size 120x112; Picture "59_1"
   GraphicView "Template_Graphic view_12" at 645,304 size 120x104; Picture "60_1"
   TextField "Template_Text field_2" at 201,80 size 20x32; Text '6'

screen "7_2" 800x480, template "Template_2"
   Button "Button_1" at 38,239 size 120x40; TextOff 'Imatinib'
      on Click: ActivateScreen("4_ORDER", 0); SetTag("Selected_URL", 'file:///C:/ASRS_Video/clip401.html')
      on Activate: SetTag("Selected_Medicine", 401)
      on Release: SetTag("ยา 401", 0)
      on Press: SetTag("ยา 401", 1)
   Button "Button_9" at 688,16 size 96x40; TextOff 'Next'
      on Press: ActivateScreen("8_2", 0)
   Button "Button_10" at 38,415 size 120x40; TextOff 'Afatinib'
      on Click: ActivateScreen("4_ORDER", 0); SetTag("Selected_URL", 'file:///C:/ASRS_Video/clip406.html')
      on Activate: SetTag("Selected_Medicine", 406)
      on Release: SetTag("ยา 406", 0)
      on Press: SetTag("ยา 406", 1)
   Button "Button_2" at 189,240 size 120x40; TextOff 'Dasatinib'
      on Click: ActivateScreen("4_ORDER", 0); SetTag("Selected_URL", 'file:///C:/ASRS_Video/clip402.html')
      on Activate: SetTag("Selected_Medicine", 402)
      on Release: SetTag("ยา 402", 0)
      on Press: SetTag("ยา 402", 1)
   Button "Button_3" at 190,415 size 120x40; TextOff 'Sunitinib'
      on Click: ActivateScreen("4_ORDER", 0); SetTag("Selected_URL", 'file:///C:/ASRS_Video/clip407.html')
      on Activate: SetTag("Selected_Medicine", 407)
      on Release: SetTag("ยา 407", 0)
      on Press: SetTag("ยา 407", 1)
   Button "Button_4" at 340,240 size 120x40; TextOff 'Nilotinib'
      on Click: ActivateScreen("4_ORDER", 0); SetTag("Selected_URL", 'file:///C:/ASRS_Video/clip403.html')
      on Activate: SetTag("Selected_Medicine", 403)
      on Release: SetTag("ยา 403", 0)
      on Press: SetTag("ยา 403", 1)
   Button "Button_5" at 340,416 size 120x40; TextOff 'Sorafenib'
      on Click: ActivateScreen("4_ORDER", 0); SetTag("Selected_URL", 'file:///C:/ASRS_Video/clip408.html')
      on Activate: SetTag("Selected_Medicine", 408)
      on Release: SetTag("ยา 408", 0)
      on Press: SetTag("ยา 408", 1)
   Button "Button_6" at 492,416 size 120x40; TextOff 'Lenvatinib'
      on Click: ActivateScreen("4_ORDER", 0); SetTag("Selected_URL", 'file:///C:/ASRS_Video/clip409.html')
      on Activate: SetTag("Selected_Medicine", 409)
      on Release: SetTag("ยา 409", 0)
      on Press: SetTag("ยา 409", 1)
   Button "Button_7" at 492,240 size 120x40; TextOff 'Erlotinib'
      on Click: ActivateScreen("4_ORDER", 0); SetTag("Selected_URL", 'file:///C:/ASRS_Video/clip404.html')
      on Activate: SetTag("Selected_Medicine", 404)
      on Release: SetTag("ยา 404", 0)
      on Press: SetTag("ยา 404", 1)
   Button "Button_8" at 644,240 size 120x40; TextOff 'Gefitinib'
      on Click: ActivateScreen("4_ORDER", 0); SetTag("Selected_URL", 'file:///C:/ASRS_Video/clip405.html')
      on Activate: SetTag("Selected_Medicine", 405)
      on Release: SetTag("ยา 405", 0)
      on Press: SetTag("ยา 405", 1)
   Button "Button_11" at 645,416 size 120x40; TextOff 'Bevacizumab'
      on Click: ActivateScreen("4_ORDER", 0); SetTag("Selected_URL", 'file:///C:/ASRS_Video/clip410.html')
      on Activate: SetTag("Selected_Medicine", 410)
      on Release: SetTag("ยา 410", 0)
      on Press: SetTag("ยา 410", 1)
   Button "Button_12" at 24,16 size 94x40; TextOff 'Back'
      on Press: ActivateScreen("6_2", 0)
   GraphicView "Template_Graphic view_1" at 693,20 size 36x32; Picture "play"
   GraphicView "Template_Graphic view_2" at 27,19 size 36x32; Picture "fast-backward"
   GraphicView "Template_Graphic view_3" at 37,128 size 120x104; Picture "61_1"
   GraphicView "Template_Graphic view_4" at 191,129 size 120x104; Picture "62_1"
   GraphicView "Template_Graphic view_5" at 339,129 size 120x104; Picture "63_1"
   GraphicView "Template_Graphic view_6" at 493,129 size 120x104; Picture "64_1"
   GraphicView "Template_Graphic view_7" at 645,129 size 120x104; Picture "65_1"
   GraphicView "Template_Graphic view_8" at 38,305 size 120x104; Picture "66_1"
   GraphicView "Template_Graphic view_9" at 189,304 size 120x112; Picture "67_1"
   GraphicView "Template_Graphic view_10" at 351,307 size 96x104; Picture "68_1"
   GraphicView "Template_Graphic view_11" at 497,304 size 120x112; Picture "69_1"
   GraphicView "Template_Graphic view_12" at 645,304 size 120x104; Picture "70_1"
   TextField "Template_Text field_2" at 201,80 size 20x32; Text '7'

screen "8_2" 800x480, template "Template_2"
   Button "Button_1" at 38,239 size 120x40; TextOff 'Trastuzumab'
      on Click: ActivateScreen("4_ORDER", 0); SetTag("Selected_URL", 'file:///C:/ASRS_Video/clip411.html')
      on Activate: SetTag("Selected_Medicine", 411)
      on Release: SetTag("ยา 411", 0)
      on Press: SetTag("ยา 411", 1)
   Button "Button_10" at 38,415 size 120x40; TextOff 'Bicalutamide'
      on Click: ActivateScreen("4_ORDER", 0); SetTag("Selected_URL", 'file:///C:/ASRS_Video/clip416.html')
      on Activate: SetTag("Selected_Medicine", 416)
      on Release: SetTag("ยา 416", 0)
      on Press: SetTag("ยา 416", 1)
   Button "Button_2" at 189,240 size 120x40; TextOff 'Rituximab'
      on Click: ActivateScreen("4_ORDER", 0); SetTag("Selected_URL", 'file:///C:/ASRS_Video/clip412.html')
      on Activate: SetTag("Selected_Medicine", 412)
      on Release: SetTag("ยา 412", 0)
      on Press: SetTag("ยา 412", 1)
   Button "Button_3" at 190,415 size 120x40; TextOff 'Flutamide'
      on Click: ActivateScreen("4_ORDER", 0); SetTag("Selected_URL", 'file:///C:/ASRS_Video/clip417.html')
      on Activate: SetTag("Selected_Medicine", 417)
      on Release: SetTag("ยา 417", 0)
      on Press: SetTag("ยา 417", 1)
   Button "Button_4" at 340,240 size 120x40; TextOff 'Pembrolizumab'
      on Click: ActivateScreen("4_ORDER", 0); SetTag("Selected_URL", 'file:///C:/ASRS_Video/clip413.html')
      on Activate: SetTag("Selected_Medicine", 413)
      on Release: SetTag("ยา 413", 0)
      on Press: SetTag("ยา 413", 1)
   Button "Button_5" at 340,416 size 120x40; TextOff 'Abiraterone'
      on Click: ActivateScreen("4_ORDER", 0); SetTag("Selected_URL", 'file:///C:/ASRS_Video/clip418.html')
      on Activate: SetTag("Selected_Medicine", 418)
      on Release: SetTag("ยา 418", 0)
      on Press: SetTag("ยา 418", 1)
   Button "Button_6" at 492,416 size 120x40; TextOff 'Enzalutamide'
      on Click: ActivateScreen("4_ORDER", 0); SetTag("Selected_URL", 'file:///C:/ASRS_Video/clip419.html')
      on Activate: SetTag("Selected_Medicine", 419)
      on Release: SetTag("ยา 419", 0)
      on Press: SetTag("ยา 419", 1)
   Button "Button_7" at 492,240 size 120x40; TextOff 'Nivolumab'
      on Click: ActivateScreen("4_ORDER", 0); SetTag("Selected_URL", 'file:///C:/ASRS_Video/clip414.html')
      on Activate: SetTag("Selected_Medicine", 414)
      on Release: SetTag("ยา 414", 0)
      on Press: SetTag("ยา 414", 1)
   Button "Button_8" at 644,240 size 120x40; TextOff 'Ipilimumab'
      on Click: ActivateScreen("4_ORDER", 0); SetTag("Selected_URL", 'file:///C:/ASRS_Video/clip415.html')
      on Activate: SetTag("Selected_Medicine", 415)
      on Release: SetTag("ยา 415", 0)
      on Press: SetTag("ยา 415", 1)
   Button "Button_11" at 645,416 size 120x40; TextOff 'Megestrol acetate'
      on Click: ActivateScreen("4_ORDER", 0); SetTag("Selected_URL", 'file:///C:/ASRS_Video/clip420.html')
      on Activate: SetTag("Selected_Medicine", 420)
      on Release: SetTag("ยา 420", 0)
      on Press: SetTag("ยา 420", 1)
   Button "Button_12" at 24,16 size 94x40; TextOff 'Back'
      on Press: ActivateScreen("7_2", 0)
   Button "Button_9" at 688,16 size 96x40; TextOff 'Next'
      on Press: ActivateScreen("9_2", 0)
   GraphicView "Template_Graphic view_2" at 27,19 size 36x32; Picture "fast-backward"
   GraphicView "Template_Graphic view_1" at 693,20 size 36x32; Picture "play"
   GraphicView "Template_Graphic view_3" at 37,128 size 120x104; Picture "71_1"
   GraphicView "Template_Graphic view_4" at 191,129 size 120x104; Picture "72_1"
   GraphicView "Template_Graphic view_5" at 339,129 size 120x104; Picture "73_1"
   GraphicView "Template_Graphic view_6" at 493,129 size 120x104; Picture "74_1"
   GraphicView "Template_Graphic view_7" at 645,129 size 120x104; Picture "75_1"
   GraphicView "Template_Graphic view_8" at 38,305 size 120x104; Picture "76_1"
   GraphicView "Template_Graphic view_9" at 189,304 size 120x112; Picture "77_1"
   GraphicView "Template_Graphic view_10" at 351,307 size 96x104; Picture "78_1"
   GraphicView "Template_Graphic view_11" at 492,303 size 120x112; Picture "79_1"
   GraphicView "Template_Graphic view_12" at 645,304 size 120x104; Picture "80_1"
   TextField "Template_Text field_2" at 201,80 size 20x32; Text '8'

screen "9_2" 800x480, template "Template_2"
   Button "Button_1" at 38,239 size 120x40; TextOff 'Zoledronic acid'
      on Click: ActivateScreen("4_ORDER", 0); SetTag("Selected_URL", 'file:///C:/ASRS_Video/clip421.html')
      on Activate: SetTag("Selected_Medicine", 421)
      on Release: SetTag("ยา 421", 0)
      on Press: SetTag("ยา 421", 1)
   Button "Button_10" at 38,415 size 120x40; TextOff 'Cyclosporine'
      on Click: ActivateScreen("4_ORDER", 0); SetTag("Selected_URL", 'file:///C:/ASRS_Video/clip426.html')
      on Activate: SetTag("Selected_Medicine", 426)
      on Release: SetTag("ยา 426", 0)
      on Press: SetTag("ยา 426", 1)
   Button "Button_2" at 189,240 size 120x40; TextOff 'Pamidronate'
      on Click: ActivateScreen("4_ORDER", 0); SetTag("Selected_URL", 'file:///C:/ASRS_Video/clip422.html')
      on Activate: SetTag("Selected_Medicine", 422)
      on Release: SetTag("ยา 422", 0)
      on Press: SetTag("ยา 422", 1)
   Button "Button_3" at 190,415 size 120x40; TextOff 'Mycophenolate mofetil'
      on Click: ActivateScreen("4_ORDER", 0); SetTag("Selected_URL", 'file:///C:/ASRS_Video/clip427.html')
      on Activate: SetTag("Selected_Medicine", 427)
      on Release: SetTag("ยา 427", 0)
      on Press: SetTag("ยา 427", 1)
   Button "Button_4" at 340,240 size 120x40; TextOff 'Calcitonin'
      on Click: ActivateScreen("4_ORDER", 0); SetTag("Selected_URL", 'file:///C:/ASRS_Video/clip423.html')
      on Activate: SetTag("Selected_Medicine", 423)
      on Release: SetTag("ยา 423", 0)
      on Press: SetTag("ยา 423", 1)
   Button "Button_5" at 340,416 size 120x40; TextOff 'Azathioprine'
      on Click: ActivateScreen("4_ORDER", 0); SetTag("Selected_URL", 'file:///C:/ASRS_Video/clip428.html')
      on Activate: SetTag("Selected_Medicine", 428)
      on Release: SetTag("ยา 428", 0)
      on Press: SetTag("ยา 428", 1)
   Button "Button_6" at 492,416 size 120x40; TextOff 'Sirolimus'
      on Click: ActivateScreen("4_ORDER", 0); SetTag("Selected_URL", 'file:///C:/ASRS_Video/clip429.html')
      on Activate: SetTag("Selected_Medicine", 429)
      on Release: SetTag("ยา 429", 0)
      on Press: SetTag("ยา 429", 1)
   Button "Button_7" at 492,240 size 120x40; TextOff 'Denosumab'
      on Click: ActivateScreen("4_ORDER", 0); SetTag("Selected_URL", 'file:///C:/ASRS_Video/clip424.html')
      on Activate: SetTag("Selected_Medicine", 424)
      on Release: SetTag("ยา 424", 0)
      on Press: SetTag("ยา 424", 1)
   Button "Button_8" at 644,240 size 120x40; TextOff 'Tacrolimus'
      on Click: ActivateScreen("4_ORDER", 0); SetTag("Selected_URL", 'file:///C:/ASRS_Video/clip425.html')
      on Activate: SetTag("Selected_Medicine", 425)
      on Release: SetTag("ยา 425", 0)
      on Press: SetTag("ยา 425", 1)
   Button "Button_11" at 645,416 size 120x40; TextOff 'Everolimus'
      on Click: ActivateScreen("4_ORDER", 0); SetTag("Selected_URL", 'file:///C:/ASRS_Video/clip430.html')
      on Activate: SetTag("Selected_Medicine", 430)
      on Release: SetTag("ยา 430", 0)
      on Press: SetTag("ยา 430", 1)
   Button "Button_12" at 24,16 size 94x40; TextOff 'Back'
      on Press: ActivateScreen("8_2", 0)
   Button "Button_9" at 688,16 size 96x40; TextOff 'Next'
      on Press: ActivateScreen("10_2", 0)
   GraphicView "Template_Graphic view_2" at 27,19 size 36x32; Picture "fast-backward"
   GraphicView "Template_Graphic view_1" at 693,20 size 36x32; Picture "play"
   GraphicView "Template_Graphic view_3" at 37,128 size 120x104; Picture "81_1"
   GraphicView "Template_Graphic view_4" at 191,129 size 120x104; Picture "82_1"
   GraphicView "Template_Graphic view_5" at 339,129 size 120x104; Picture "83_1"
   GraphicView "Template_Graphic view_6" at 493,129 size 120x104; Picture "84_1"
   GraphicView "Template_Graphic view_7" at 645,129 size 120x104; Picture "85_1"
   GraphicView "Template_Graphic view_8" at 38,305 size 120x104; Picture "86_1"
   GraphicView "Template_Graphic view_9" at 189,304 size 120x112; Picture "87_1"
   GraphicView "Template_Graphic view_10" at 351,307 size 96x104; Picture "88_1"
   GraphicView "Template_Graphic view_11" at 497,304 size 120x112; Picture "89_1"
   GraphicView "Template_Graphic view_12" at 645,304 size 120x104; Picture "90_1"
   TextField "Template_Text field_2" at 201,80 size 20x32; Text '9'

screen "10_2" 800x480, template "Template_2"
   Button "Button_1" at 38,239 size 120x40; TextOff 'Prednisolone'
      on Click: ActivateScreen("4_ORDER", 0); SetTag("Selected_URL", 'file:///C:/ASRS_Video/clip431.html')
      on Activate: SetTag("Selected_Medicine", 431)
      on Release: SetTag("ยา 431", 0)
      on Press: SetTag("ยา 431", 1)
   Button "Button_10" at 38,415 size 120x40; TextOff 'Interferon alfa'
      on Click: ActivateScreen("4_ORDER", 0); SetTag("Selected_URL", 'file:///C:/ASRS_Video/clip436.html')
      on Activate: SetTag("Selected_Medicine", 436)
      on Release: SetTag("ยา 436", 0)
      on Press: SetTag("ยา 436", 1)
   Button "Button_2" at 189,240 size 120x40; TextOff 'Methylprednisolone'
      on Click: ActivateScreen("4_ORDER", 0); SetTag("Selected_URL", 'file:///C:/ASRS_Video/clip432.html')
      on Activate: SetTag("Selected_Medicine", 432)
      on Release: SetTag("ยา 432", 0)
      on Press: SetTag("ยา 432", 1)
   Button "Button_3" at 190,415 size 120x40; TextOff 'Epoetin alfa'
      on Click: ActivateScreen("4_ORDER", 0); SetTag("Selected_URL", 'file:///C:/ASRS_Video/clip437.html')
      on Activate: SetTag("Selected_Medicine", 437)
      on Release: SetTag("ยา 437", 0)
      on Press: SetTag("ยา 437", 1)
   Button "Button_4" at 340,240 size 120x40; TextOff 'Dexamethasone'
      on Click: ActivateScreen("4_ORDER", 0); SetTag("Selected_URL", 'file:///C:/ASRS_Video/clip433.html')
      on Activate: SetTag("Selected_Medicine", 433)
      on Release: SetTag("ยา 433", 0)
      on Press: SetTag("ยา 433", 1)
   Button "Button_5" at 340,416 size 120x40; TextOff 'Filgrastim'
      on Click: ActivateScreen("4_ORDER", 0); SetTag("Selected_URL", 'file:///C:/ASRS_Video/clip438.html')
      on Activate: SetTag("Selected_Medicine", 438)
      on Release: SetTag("ยา 438", 0)
      on Press: SetTag("ยา 438", 1)
   Button "Button_6" at 492,416 size 120x40; TextOff 'Pegfilgrastim'
      on Click: ActivateScreen("4_ORDER", 0); SetTag("Selected_URL", 'file:///C:/ASRS_Video/clip439.html')
      on Activate: SetTag("Selected_Medicine", 439)
      on Release: SetTag("ยา 439", 0)
      on Press: SetTag("ยา 439", 1)
   Button "Button_7" at 492,240 size 120x40; TextOff 'Basiliximab'
      on Click: ActivateScreen("4_ORDER", 0); SetTag("Selected_URL", 'file:///C:/ASRS_Video/clip434.html')
      on Activate: SetTag("Selected_Medicine", 434)
      on Release: SetTag("ยา 434", 0)
      on Press: SetTag("ยา 434", 1)
   Button "Button_8" at 644,240 size 120x40; TextOff 'Anti-thymocyte globulin'
      on Click: ActivateScreen("4_ORDER", 0); SetTag("Selected_URL", 'file:///C:/ASRS_Video/clip435.html')
      on Activate: SetTag("Selected_Medicine", 435)
      on Release: SetTag("ยา 435", 0)
      on Press: SetTag("ยา 435", 1)
   Button "Button_11" at 645,416 size 120x40; TextOff 'Romiplostim'
      on Click: ActivateScreen("4_ORDER", 0); SetTag("Selected_URL", 'file:///C:/ASRS_Video/clip440.html')
      on Activate: SetTag("Selected_Medicine", 440)
      on Release: SetTag("ยา 440", 0)
      on Press: SetTag("ยา 440", 1)
   Button "Button_12" at 24,16 size 94x40; TextOff 'Back'
      on Press: ActivateScreen("9_2", 0)
   Button "Button_9" at 688,16 size 96x40; TextOff 'Next'
      on Press: ActivateScreen("11_2", 0)
   GraphicView "Template_Graphic view_2" at 27,19 size 36x32; Picture "fast-backward"
   GraphicView "Template_Graphic view_1" at 693,20 size 36x32; Picture "play"
   GraphicView "Template_Graphic view_3" at 37,128 size 120x104; Picture "91_1"
   GraphicView "Template_Graphic view_4" at 191,129 size 120x104; Picture "92_1"
   GraphicView "Template_Graphic view_5" at 339,129 size 120x104; Picture "93_1"
   GraphicView "Template_Graphic view_6" at 493,129 size 120x104; Picture "94_1"
   GraphicView "Template_Graphic view_7" at 645,129 size 120x104; Picture "95_1"
   GraphicView "Template_Graphic view_8" at 38,305 size 120x104; Picture "96_1"
   GraphicView "Template_Graphic view_9" at 189,304 size 120x112; Picture "97_1"
   GraphicView "Template_Graphic view_10" at 351,307 size 96x104; Picture "98_1"
   GraphicView "Template_Graphic view_11" at 497,304 size 120x112; Picture "99_1"
   GraphicView "Template_Graphic view_12" at 645,304 size 120x104; Picture "100_1"
   TextField "Template_Text field_2" at 201,80 size 36x32; Text '10'

screen "11_2" 800x480, template "Template_2"
   Button "Button_1" at 38,239 size 120x40; TextOff 'Thalidomide'
      on Click: ActivateScreen("4_ORDER", 0); SetTag("Selected_URL", 'file:///C:/ASRS_Video/clip441.html')
      on Activate: SetTag("Selected_Medicine", 441)
      on Release: SetTag("ยา 441", 0)
      on Press: SetTag("ยา 441", 1)
   Button "Button_10" at 38,415 size 120x40; TextOff 'Mesna'
      on Click: ActivateScreen("4_ORDER", 0); SetTag("Selected_URL", 'file:///C:/ASRS_Video/clip446.html')
      on Activate: SetTag("Selected_Medicine", 446)
      on Release: SetTag("ยา 446", 0)
      on Press: SetTag("ยา 446", 1)
   Button "Button_2" at 189,240 size 120x40; TextOff 'Lenalidomide'
      on Click: ActivateScreen("4_ORDER", 0); SetTag("Selected_URL", 'file:///C:/ASRS_Video/clip442.html')
      on Activate: SetTag("Selected_Medicine", 442)
      on Release: SetTag("ยา 442", 0)
      on Press: SetTag("ยา 442", 1)
   Button "Button_3" at 190,415 size 120x40; TextOff 'Leucovorin'
      on Click: ActivateScreen("4_ORDER", 0); SetTag("Selected_URL", 'file:///C:/ASRS_Video/clip447.html')
      on Activate: SetTag("Selected_Medicine", 447)
      on Release: SetTag("ยา 447", 0)
      on Press: SetTag("ยา 447", 1)
   Button "Button_4" at 340,240 size 120x40; TextOff 'Bortezomib'
      on Click: ActivateScreen("4_ORDER", 0); SetTag("Selected_URL", 'file:///C:/ASRS_Video/clip443.html')
      on Activate: SetTag("Selected_Medicine", 443)
      on Release: SetTag("ยา 443", 0)
      on Press: SetTag("ยา 443", 1)
   Button "Button_5" at 340,416 size 120x40; TextOff 'All-trans retinoic acid'
      on Click: ActivateScreen("4_ORDER", 0); SetTag("Selected_URL", 'file:///C:/ASRS_Video/clip448.html')
      on Activate: SetTag("Selected_Medicine", 448)
      on Release: SetTag("ยา 448", 0)
      on Press: SetTag("ยา 448", 1)
   Button "Button_6" at 492,416 size 120x40; TextOff 'Arsenic trioxide'
      on Click: ActivateScreen("4_ORDER", 0); SetTag("Selected_URL", 'file:///C:/ASRS_Video/clip449.html')
      on Activate: SetTag("Selected_Medicine", 449)
      on Release: SetTag("ยา 449", 0)
      on Press: SetTag("ยา 449", 1)
   Button "Button_7" at 492,240 size 120x40; TextOff 'Carfilzomib'
      on Click: ActivateScreen("4_ORDER", 0); SetTag("Selected_URL", 'file:///C:/ASRS_Video/clip444.html')
      on Activate: SetTag("Selected_Medicine", 444)
      on Release: SetTag("ยา 444", 0)
      on Press: SetTag("ยา 444", 1)
   Button "Button_8" at 644,240 size 120x40; TextOff 'Daratumumab'
      on Click: ActivateScreen("4_ORDER", 0); SetTag("Selected_URL", 'file:///C:/ASRS_Video/clip445.html')
      on Activate: SetTag("Selected_Medicine", 445)
      on Release: SetTag("ยา 445", 0)
      on Press: SetTag("ยา 445", 1)
   Button "Button_11" at 645,416 size 120x40; TextOff 'Temozolomide'
      on Click: ActivateScreen("4_ORDER", 0); SetTag("Selected_URL", 'file:///C:/ASRS_Video/clip450.html')
      on Activate: SetTag("Selected_Medicine", 450)
      on Release: SetTag("ยา 450", 0)
      on Press: SetTag("ยา 450", 1)
   Button "Button_12" at 24,16 size 94x40; TextOff 'Back'
      on Press: ActivateScreen("10_2", 0)
   Button "Button_9" at 688,16 size 96x40; TextOff 'Next'
      on Press: ActivateScreen("12_2", 0)
   GraphicView "Template_Graphic view_2" at 27,19 size 36x32; Picture "fast-backward"
   GraphicView "Template_Graphic view_1" at 693,20 size 36x32; Picture "play"
   GraphicView "Template_Graphic view_3" at 37,128 size 120x104; Picture "101_1"
   GraphicView "Template_Graphic view_4" at 191,129 size 120x104; Picture "102_1"
   GraphicView "Template_Graphic view_5" at 339,129 size 120x104; Picture "103_1"
   GraphicView "Template_Graphic view_6" at 493,129 size 120x104; Picture "104_1"
   GraphicView "Template_Graphic view_7" at 645,129 size 120x104; Picture "105_1"
   GraphicView "Template_Graphic view_8" at 38,305 size 120x104; Picture "106_1"
   GraphicView "Template_Graphic view_9" at 189,304 size 120x112; Picture "107_1"
   GraphicView "Template_Graphic view_10" at 351,307 size 96x104; Picture "108_1"
   GraphicView "Template_Graphic view_11" at 497,304 size 120x112; Picture "109_1"
   GraphicView "Template_Graphic view_12" at 645,304 size 120x104; Picture "110_1"
   TextField "Template_Text field_2" at 201,80 size 36x32; Text '11'

screen "12_2" 800x480, template "Template_2"
   Button "Button_1" at 38,239 size 120x40; TextOff 'Procarbazine'
      on Click: ActivateScreen("4_ORDER", 0); SetTag("Selected_URL", 'file:///C:/ASRS_Video/clip451.html')
      on Activate: SetTag("Selected_Medicine", 451)
      on Release: SetTag("ยา 451", 0)
      on Press: SetTag("ยา 451", 1)
   Button "Button_10" at 38,415 size 120x40; TextOff 'Asparaginase'
      on Click: ActivateScreen("4_ORDER", 0); SetTag("Selected_URL", 'file:///C:/ASRS_Video/clip456.html')
      on Activate: SetTag("Selected_Medicine", 456)
      on Release: SetTag("ยา 456", 0)
      on Press: SetTag("ยา 456", 1)
   Button "Button_2" at 189,240 size 120x40; TextOff 'Lomustine'
      on Click: ActivateScreen("4_ORDER", 0); SetTag("Selected_URL", 'file:///C:/ASRS_Video/clip452.html')
      on Activate: SetTag("Selected_Medicine", 452)
      on Release: SetTag("ยา 452", 0)
      on Press: SetTag("ยา 452", 1)
   Button "Button_3" at 190,415 size 120x40; TextOff 'Pegaspargase'
      on Click: ActivateScreen("4_ORDER", 0); SetTag("Selected_URL", 'file:///C:/ASRS_Video/clip457.html')
      on Activate: SetTag("Selected_Medicine", 457)
      on Release: SetTag("ยา 457", 0)
      on Press: SetTag("ยา 457", 1)
   Button "Button_4" at 340,240 size 120x40; TextOff 'Carmustine'
      on Click: ActivateScreen("4_ORDER", 0); SetTag("Selected_URL", 'file:///C:/ASRS_Video/clip453.html')
      on Activate: SetTag("Selected_Medicine", 453)
      on Release: SetTag("ยา 453", 0)
      on Press: SetTag("ยา 453", 1)
   Button "Button_5" at 340,416 size 120x40; TextOff 'Brentuximab vedotin'
      on Click: ActivateScreen("4_ORDER", 0); SetTag("Selected_URL", 'file:///C:/ASRS_Video/clip458.html')
      on Activate: SetTag("Selected_Medicine", 458)
      on Release: SetTag("ยา 458", 0)
      on Press: SetTag("ยา 458", 1)
   Button "Button_6" at 492,416 size 120x40; TextOff 'Olaparib'
      on Click: ActivateScreen("4_ORDER", 0); SetTag("Selected_URL", 'file:///C:/ASRS_Video/clip459.html')
      on Activate: SetTag("Selected_Medicine", 459)
      on Release: SetTag("ยา 459", 0)
      on Press: SetTag("ยา 459", 1)
   Button "Button_7" at 492,240 size 120x40; TextOff 'Mitomycin C'
      on Click: ActivateScreen("4_ORDER", 0); SetTag("Selected_URL", 'file:///C:/ASRS_Video/clip454.html')
      on Activate: SetTag("Selected_Medicine", 454)
      on Release: SetTag("ยา 454", 0)
      on Press: SetTag("ยา 454", 1)
   Button "Button_8" at 644,240 size 120x40; TextOff 'Actinomycin D'
      on Click: ActivateScreen("4_ORDER", 0); SetTag("Selected_URL", 'file:///C:/ASRS_Video/clip455.html')
      on Activate: SetTag("Selected_Medicine", 455)
      on Release: SetTag("ยา 455", 0)
      on Press: SetTag("ยา 455", 1)
   Button "Button_11" at 645,416 size 120x40; TextOff 'Palbociclib'
      on Click: ActivateScreen("4_ORDER", 0); SetTag("Selected_URL", 'file:///C:/ASRS_Video/clip460.html')
      on Activate: SetTag("Selected_Medicine", 460)
      on Release: SetTag("ยา 460", 0)
      on Press: SetTag("ยา 460", 1)
   Button "Button_12" at 24,16 size 94x40; TextOff 'Back'
      on Press: ActivateScreen("11_2", 0)
   GraphicView "Template_Graphic view_2" at 27,19 size 36x32; Picture "fast-backward"
   GraphicView "Template_Graphic view_3" at 37,128 size 120x104; Picture "111_1"
   GraphicView "Template_Graphic view_4" at 191,129 size 120x104; Picture "112_1"
   GraphicView "Template_Graphic view_5" at 339,129 size 120x104; Picture "113_1"
   GraphicView "Template_Graphic view_6" at 493,129 size 120x104; Picture "114_1"
   GraphicView "Template_Graphic view_7" at 645,129 size 120x104; Picture "115_1"
   GraphicView "Template_Graphic view_8" at 38,305 size 120x104; Picture "116_1"
   GraphicView "Template_Graphic view_9" at 189,304 size 120x112; Picture "117_1"
   GraphicView "Template_Graphic view_10" at 351,307 size 96x104; Picture "118_1"
   GraphicView "Template_Graphic view_11" at 497,304 size 120x112; Picture "119_1"
   GraphicView "Template_Graphic view_12" at 645,304 size 120x104; Picture "120_1"
   TextField "Template_Text field_2" at 201,80 size 36x32; Text '12'

screen "1_1" 800x480, template "Template_2"
   Button "Button_1" at 40,240 size 120x40; TextOff 'Amoxicillin'
      on Click: ActivateScreen("4_ORDER", 0); SetTag("Selected_URL", 'file:///C:/ASRS_Video/clip221.html')
      on Activate: SetTag("Selected_Medicine", 221)
      on Release: SetTag("ยา 221", 0)
      on Press: SetTag("ยา 221", 1)
   Button "Button_10" at 38,415 size 120x40; TextOff 'Benzathine penicillin G'
      on Click: ActivateScreen("4_ORDER", 0); SetTag("Selected_URL", 'file:///C:/ASRS_Video/clip226.html')
      on Activate: SetTag("Selected_Medicine", 227)
      on Release: SetTag("ยา 226", 0)
      on Press: SetTag("ยา 226", 1)
   Button "Button_2" at 189,240 size 120x40; TextOff 'Ampicillin'
      on Click: ActivateScreen("4_ORDER", 0); SetTag("Selected_URL", 'file:///C:/ASRS_Video/clip222.html')
      on Activate: SetTag("Selected_Medicine", 222)
      on Release: SetTag("ยา 222", 0)
      on Press: SetTag("ยา 222", 1)
   Button "Button_3" at 190,415 size 120x40; TextOff 'Piperacillin'
      on Click: ActivateScreen("4_ORDER", 0); SetTag("Selected_URL", 'file:///C:/ASRS_Video/clip227.html')
      on Activate: SetTag("Selected_Medicine", 228)
      on Release: SetTag("ยา 227", 0)
      on Press: SetTag("ยา 227", 1)
   Button "Button_4" at 340,240 size 120x40; TextOff 'Cloxacillin'
      on Click: ActivateScreen("4_ORDER", 0); SetTag("Selected_URL", 'file:///C:/ASRS_Video/clip223.html')
      on Activate: SetTag("Selected_Medicine", 223)
      on Release: SetTag("ยา 223", 0)
      on Press: SetTag("ยา 223", 1)
   Button "Button_5" at 340,416 size 120x40; TextOff 'Ticarcillin'
      on Click: ActivateScreen("4_ORDER", 0); SetTag("Selected_URL", 'file:///C:/ASRS_Video/clip228.html')
      on Activate: SetTag("Selected_Medicine", 229)
      on Release: SetTag("ยา 228", 0)
      on Press: SetTag("ยา 228", 1)
   Button "Button_6" at 492,416 size 120x40; TextOff 'Amoxicillin clavulanate'
      on Click: ActivateScreen("4_ORDER", 0); SetTag("Selected_URL", 'file:///C:/ASRS_Video/clip229.html')
      on Activate: SetTag("Selected_Medicine", 230)
      on Release: SetTag("ยา 229", 0)
      on Press: SetTag("ยา 229", 1)
   Button "Button_7" at 492,240 size 120x40; TextOff 'Dicloxacillin'
      on Click: ActivateScreen("4_ORDER", 0); SetTag("Selected_URL", 'file:///C:/ASRS_Video/clip224.html')
      on Activate: SetTag("Selected_Medicine", 224)
      on Release: SetTag("ยา 224", 0)
      on Press: SetTag("ยา 224", 1)
   Button "Button_8" at 644,240 size 120x40; TextOff 'Penicillin V'
      on Click: ActivateScreen("4_ORDER", 0); SetTag("Selected_URL", 'file:///C:/ASRS_Video/clip225.html')
      on Activate: SetTag("Selected_Medicine", 225)
      on Release: SetTag("ยา 225", 0)
      on Press: SetTag("ยา 225", 1)
   Button "Button_11" at 645,416 size 120x40; TextOff 'Ampicillin sulbactam'
      on Click: ActivateScreen("4_ORDER", 0); SetTag("Selected_URL", 'file:///C:/ASRS_Video/clip230.html')
      on Activate: SetTag("Selected_Medicine", 230)
      on Release: SetTag("ยา 230", 0)
      on Press: SetTag("ยา 230", 1)
   Button "Button_12" at 688,16 size 96x40; TextOff 'Next'
      on Press: ActivateScreen("2_1", 0)
   Button "Button_9" at 24,16 size 94x40; TextOff 'Back'
      on Press: ActivateScreen("4_ORDER", 0)
   GraphicView "Template_Graphic view_2" at 693,20 size 36x32; Picture "play"
   GraphicView "Template_Graphic view_1" at 27,19 size 36x32; Picture "fast-backward"
   GraphicView "Template_Graphic view_3" at 37,128 size 120x104; Picture "1"
   GraphicView "Template_Graphic view_4" at 191,129 size 120x104; Picture "2"
   GraphicView "Template_Graphic view_5" at 339,129 size 120x104; Picture "3"
   GraphicView "Template_Graphic view_6" at 493,129 size 120x104; Picture "4"
   GraphicView "Template_Graphic view_7" at 645,129 size 120x104; Picture "5"
   GraphicView "Template_Graphic view_8" at 38,305 size 120x104; Picture "6"
   GraphicView "Template_Graphic view_9" at 189,304 size 120x112; Picture "7"
   GraphicView "Template_Graphic view_10" at 351,307 size 96x104; Picture "8"
   GraphicView "Template_Graphic view_11" at 497,304 size 120x112; Picture "9"
   GraphicView "Template_Graphic view_12" at 645,304 size 120x104; Picture "10"
   TextField "Template_Text field_2" at 201,80 size 20x32; Text '1'

screen "2_1" 800x480, template "Template_2"
   Button "Button_1" at 40,240 size 120x40; TextOff 'Cefalexin'
      on Click: ActivateScreen("4_ORDER", 0); SetTag("Selected_URL", 'file:///C:/ASRS_Video/clip231.html')
      on Activate: SetTag("Selected_Medicine", 231)
      on Release: SetTag("ยา 231", 0)
      on Press: SetTag("ยา 231", 1)
   Button "Button_9" at 688,16 size 96x40; TextOff 'Next'
      on Press: ActivateScreen("3_1", 0)
   Button "Button_10" at 40,416 size 120x40; TextOff 'Ceftriaxone'
      on Click: ActivateScreen("4_ORDER", 0); SetTag("Selected_URL", 'file:///C:/ASRS_Video/clip236.html')
      on Activate: SetTag("Selected_Medicine", 236)
      on Release: SetTag("ยา 236", 0)
      on Press: SetTag("ยา 236", 1)
   Button "Button_2" at 191,241 size 120x40; TextOff 'Cefadroxil'
      on Click: ActivateScreen("4_ORDER", 0); SetTag("Selected_URL", 'file:///C:/ASRS_Video/clip232.html')
      on Activate: SetTag("Selected_Medicine", 232)
      on Release: SetTag("ยา 232", 0)
      on Press: SetTag("ยา 232", 1)
   Button "Button_3" at 192,416 size 120x40; TextOff 'Cefotaxime'
      on Click: ActivateScreen("4_ORDER", 0); SetTag("Selected_URL", 'file:///C:/ASRS_Video/clip237.html')
      on Activate: SetTag("Selected_Medicine", 237)
      on Release: SetTag("ยา 237", 0)
      on Press: SetTag("ยา 237", 1)
   Button "Button_4" at 342,241 size 120x40; TextOff 'Cefuroxime'
      on Click: ActivateScreen("4_ORDER", 0); SetTag("Selected_URL", 'file:///C:/ASRS_Video/clip233.html')
      on Activate: SetTag("Selected_Medicine", 233)
      on Release: SetTag("ยา 233", 0)
      on Press: SetTag("ยา 233", 1)
   Button "Button_5" at 340,416 size 120x40; TextOff 'Ceftazidime'
      on Click: ActivateScreen("4_ORDER", 0); SetTag("Selected_URL", 'file:///C:/ASRS_Video/clip238.html')
      on Activate: SetTag("Selected_Medicine", 238)
      on Release: SetTag("ยา 238", 0)
      on Press: SetTag("ยา 238", 1)
   Button "Button_6" at 492,416 size 120x40; TextOff 'Cefepime'
      on Click: ActivateScreen("4_ORDER", 0); SetTag("Selected_URL", 'file:///C:/ASRS_Video/clip239.html')
      on Activate: SetTag("Selected_Medicine", 289)
      on Release: SetTag("ยา 239", 0)
      on Press: SetTag("ยา 239", 1)
   Button "Button_7" at 492,240 size 120x40; TextOff 'Cefixime'
      on Click: ActivateScreen("4_ORDER", 0); SetTag("Selected_URL", 'file:///C:/ASRS_Video/clip234.html')
      on Activate: SetTag("Selected_Medicine", 234)
      on Release: SetTag("ยา 234", 0)
      on Press: SetTag("ยา 234", 1)
   Button "Button_8" at 644,240 size 120x40; TextOff 'Cefpodoxime'
      on Click: ActivateScreen("4_ORDER", 0); SetTag("Selected_URL", 'file:///C:/ASRS_Video/clip235.html')
      on Activate: SetTag("Selected_Medicine", 235)
      on Release: SetTag("ยา 235", 0)
      on Press: SetTag("ยา 235", 1)
   Button "Button_11" at 645,416 size 120x40; TextOff 'Cefoxitin'
      on Click: ActivateScreen("4_ORDER", 0); SetTag("Selected_URL", 'file:///C:/ASRS_Video/clip240.html')
      on Activate: SetTag("Selected_Medicine", 240)
      on Release: SetTag("ยา 240", 0)
      on Press: SetTag("ยา 240", 1)
   Button "Button_12" at 24,16 size 94x40; TextOff 'Back'
      on Press: ActivateScreen("1_1", 0)
   GraphicView "Template_Graphic view_1" at 693,20 size 36x32; Picture "play"
   GraphicView "Template_Graphic view_2" at 27,19 size 36x32; Picture "fast-backward"
   GraphicView "Template_Graphic view_3" at 37,128 size 120x104; Picture "11"
   GraphicView "Template_Graphic view_4" at 191,129 size 120x104; Picture "12"
   GraphicView "Template_Graphic view_5" at 339,129 size 120x104; Picture "13"
   GraphicView "Template_Graphic view_6" at 493,129 size 120x104; Picture "14"
   GraphicView "Template_Graphic view_7" at 645,129 size 120x104; Picture "15"
   GraphicView "Template_Graphic view_8" at 38,305 size 120x104; Picture "16"
   GraphicView "Template_Graphic view_9" at 189,304 size 120x112; Picture "17"
   GraphicView "Template_Graphic view_10" at 351,307 size 96x104; Picture "18"
   GraphicView "Template_Graphic view_11" at 497,304 size 120x112; Picture "19"
   GraphicView "Template_Graphic view_12" at 645,304 size 120x104; Picture "20"
   TextField "Template_Text field_2" at 201,80 size 20x32; Text '2'

screen "3_1" 800x480, template "Template_2"
   Button "Button_1" at 38,239 size 120x40; TextOff 'Imipenem cilastatin'
      on Click: ActivateScreen("4_ORDER", 0); SetTag("Selected_URL", 'file:///C:/ASRS_Video/clip241.html')
      on Activate: SetTag("Selected_Medicine", 241)
      on Release: SetTag("ยา 241", 0)
      on Press: SetTag("ยา 241", 1)
   Button "Button_9" at 688,16 size 96x40; TextOff 'Next'
      on Press: ActivateScreen("4_1", 0)
   Button "Button_10" at 38,415 size 120x40; TextOff 'Teicoplanin'
      on Click: ActivateScreen("4_ORDER", 0); SetTag("Selected_URL", 'file:///C:/ASRS_Video/clip246.html')
      on Activate: SetTag("Selected_Medicine", 246)
      on Release: SetTag("ยา 246", 0)
      on Press: SetTag("ยา 246", 1)
   Button "Button_2" at 189,240 size 120x40; TextOff 'Meropenem'
      on Click: ActivateScreen("4_ORDER", 0); SetTag("Selected_URL", 'file:///C:/ASRS_Video/clip242.html')
      on Activate: SetTag("Selected_Medicine", 242)
      on Release: SetTag("ยา 242", 0)
      on Press: SetTag("ยา 242", 1)
   Button "Button_3" at 190,415 size 120x40; TextOff 'Linezolid'
      on Click: ActivateScreen("4_ORDER", 0); SetTag("Selected_URL", 'file:///C:/ASRS_Video/clip247.html')
      on Activate: SetTag("Selected_Medicine", 247)
      on Release: SetTag("ยา 246", 0)
      on Press: SetTag("ยา 247", 1)
   Button "Button_4" at 340,240 size 120x40; TextOff 'Ertapenem'
      on Click: ActivateScreen("4_ORDER", 0); SetTag("Selected_URL", 'file:///C:/ASRS_Video/clip243.html')
      on Activate: SetTag("Selected_Medicine", 243)
      on Release: SetTag("ยา 243", 0)
      on Press: SetTag("ยา 243", 1)
   Button "Button_5" at 340,416 size 120x40; TextOff 'Daptomycin'
      on Click: ActivateScreen("4_ORDER", 0); SetTag("Selected_URL", 'file:///C:/ASRS_Video/clip248.html')
      on Activate: SetTag("Selected_Medicine", 248)
      on Release: SetTag("ยา 248", 0)
      on Press: SetTag("ยา 248", 1)
   Button "Button_6" at 492,416 size 120x40; TextOff 'Gentamicin'
      on Click: ActivateScreen("4_ORDER", 0); SetTag("Selected_URL", 'file:///C:/ASRS_Video/clip249.html')
      on Activate: SetTag("Selected_Medicine", 249)
      on Release: SetTag("ยา 249", 0)
      on Press: SetTag("ยา 249", 1)
   Button "Button_7" at 492,240 size 120x40; TextOff 'Aztreonam'
      on Click: ActivateScreen("4_ORDER", 0); SetTag("Selected_URL", 'file:///C:/ASRS_Video/clip244.html')
      on Activate: SetTag("Selected_Medicine", 244)
      on Release: SetTag("ยา 244", 0)
      on Press: SetTag("ยา 244", 1)
   Button "Button_8" at 644,240 size 120x40; TextOff 'Vancomycin'
      on Click: ActivateScreen("4_ORDER", 0); SetTag("Selected_URL", 'file:///C:/ASRS_Video/clip245.html')
      on Activate: SetTag("Selected_Medicine", 245)
      on Release: SetTag("ยา 245", 0)
      on Press: SetTag("ยา 245", 1)
   Button "Button_11" at 645,416 size 120x40; TextOff 'Amikacin'
      on Click: ActivateScreen("4_ORDER", 0); SetTag("Selected_URL", 'file:///C:/ASRS_Video/clip250.html')
      on Activate: SetTag("Selected_Medicine", 250)
      on Release: SetTag("ยา 250", 0)
      on Press: SetTag("ยา 250", 1)
   Button "Button_12" at 24,16 size 94x40; TextOff 'Back'
      on Press: ActivateScreen("2_1", 0)
   GraphicView "Template_Graphic view_1" at 693,20 size 36x32; Picture "play"
   GraphicView "Template_Graphic view_2" at 27,19 size 36x32; Picture "fast-backward"
   GraphicView "Template_Graphic view_3" at 37,128 size 120x104; Picture "21"
   GraphicView "Template_Graphic view_4" at 191,129 size 120x104; Picture "22"
   GraphicView "Template_Graphic view_5" at 339,129 size 120x104; Picture "23"
   GraphicView "Template_Graphic view_6" at 493,129 size 120x104; Picture "24"
   GraphicView "Template_Graphic view_7" at 645,129 size 120x104; Picture "25"
   GraphicView "Template_Graphic view_8" at 38,305 size 120x104; Picture "26"
   GraphicView "Template_Graphic view_9" at 189,304 size 120x112; Picture "27"
   GraphicView "Template_Graphic view_10" at 351,307 size 96x104; Picture "28"
   GraphicView "Template_Graphic view_11" at 497,304 size 120x112; Picture "29"
   GraphicView "Template_Graphic view_12" at 645,304 size 120x104; Picture "30"
   TextField "Template_Text field_2" at 201,80 size 20x32; Text '3'

screen "4_1" 800x480, template "Template_2"
   Button "Button_1" at 38,239 size 120x40; TextOff 'Tobramycin'
      on Click: ActivateScreen("4_ORDER", 0); SetTag("Selected_URL", 'file:///C:/ASRS_Video/clip251.html')
      on Activate: SetTag("Selected_Medicine", 251)
      on Release: SetTag("ยา 251", 0)
      on Press: SetTag("ยา 251", 1)
   Button "Button_9" at 688,16 size 96x40; TextOff 'Next'
      on Press: ActivateScreen("5_1", 0)
   Button "Button_10" at 38,415 size 120x40; TextOff 'Azithromycin'
      on Click: ActivateScreen("4_ORDER", 0); SetTag("Selected_URL", 'file:///C:/ASRS_Video/clip256.html')
      on Activate: SetTag("Selected_Medicine", 256)
      on Release: SetTag("ยา 256", 0)
      on Press: SetTag("ยา 256", 1)
   Button "Button_2" at 189,240 size 120x40; TextOff 'Streptomycin'
      on Click: ActivateScreen("4_ORDER", 0); SetTag("Selected_URL", 'file:///C:/ASRS_Video/clip252.html')
      on Activate: SetTag("Selected_Medicine", 252)
      on Release: SetTag("ยา 252", 0)
      on Press: SetTag("ยา 252", 1)
   Button "Button_3" at 190,415 size 120x40; TextOff 'Roxithromycin'
      on Click: ActivateScreen("4_ORDER", 0); SetTag("Selected_URL", 'file:///C:/ASRS_Video/clip257.html')
      on Activate: SetTag("Selected_Medicine", 257)
      on Release: SetTag("ยา 257", 0)
      on Press: SetTag("ยา 257", 1)
   Button "Button_4" at 340,240 size 120x40; TextOff 'Neomycin'
      on Click: ActivateScreen("4_ORDER", 0); SetTag("Selected_URL", 'file:///C:/ASRS_Video/clip253.html')
      on Activate: SetTag("Selected_Medicine", 253)
      on Release: SetTag("ยา 253", 0)
      on Press: SetTag("ยา 253", 1)
   Button "Button_5" at 340,416 size 120x40; TextOff 'Clindamycin'
      on Click: ActivateScreen("4_ORDER", 0); SetTag("Selected_URL", 'file:///C:/ASRS_Video/clip258.html')
      on Activate: SetTag("Selected_Medicine", 258)
      on Release: SetTag("ยา 258", 0)
      on Press: SetTag("ยา 258", 1)
   Button "Button_6" at 492,416 size 120x40; TextOff 'Lincomycin'
      on Click: ActivateScreen("4_ORDER", 0); SetTag("Selected_URL", 'file:///C:/ASRS_Video/clip259.html')
      on Activate: SetTag("Selected_Medicine", 259)
      on Release: SetTag("ยา 259", 0)
      on Press: SetTag("ยา 259", 1)
   Button "Button_7" at 492,240 size 120x40; TextOff 'Erythromycin'
      on Click: ActivateScreen("4_ORDER", 0); SetTag("Selected_URL", 'file:///C:/ASRS_Video/clip254.html')
      on Activate: SetTag("Selected_Medicine", 254)
      on Release: SetTag("ยา 254", 0)
      on Press: SetTag("ยา 254", 1)
   Button "Button_8" at 644,240 size 120x40; TextOff 'Clarithromycin'
      on Click: ActivateScreen("4_ORDER", 0); SetTag("Selected_URL", 'file:///C:/ASRS_Video/clip255.html')
      on Activate: SetTag("Selected_Medicine", 255)
      on Release: SetTag("ยา 255", 0)
      on Press: SetTag("ยา 255", 1)
   Button "Button_11" at 645,416 size 120x40; TextOff 'Doxycycline'
      on Click: ActivateScreen("4_ORDER", 0); SetTag("Selected_URL", 'file:///C:/ASRS_Video/clip260.html')
      on Activate: SetTag("Selected_Medicine", 260)
      on Release: SetTag("ยา 260", 0)
      on Press: SetTag("ยา 260", 1)
   Button "Button_12" at 24,16 size 94x40; TextOff 'Back'
      on Press: ActivateScreen("3_1", 0)
   GraphicView "Template_Graphic view_1" at 693,20 size 36x32; Picture "play"
   GraphicView "Template_Graphic view_2" at 27,19 size 36x32; Picture "fast-backward"
   GraphicView "Template_Graphic view_3" at 37,128 size 120x104; Picture "31"
   GraphicView "Template_Graphic view_4" at 191,129 size 120x104; Picture "32"
   GraphicView "Template_Graphic view_5" at 339,129 size 120x104; Picture "33"
   GraphicView "Template_Graphic view_6" at 493,129 size 120x104; Picture "34"
   GraphicView "Template_Graphic view_7" at 645,129 size 120x104; Picture "35"
   GraphicView "Template_Graphic view_8" at 38,305 size 120x104; Picture "36"
   GraphicView "Template_Graphic view_9" at 189,304 size 120x112; Picture "37"
   GraphicView "Template_Graphic view_10" at 351,307 size 96x104; Picture "38"
   GraphicView "Template_Graphic view_11" at 497,304 size 120x112; Picture "39"
   GraphicView "Template_Graphic view_12" at 645,304 size 120x104; Picture "40"
   TextField "Template_Text field_2" at 201,80 size 20x32; Text '4'

screen "5_1" 800x480, template "Template_2"
   Button "Button_1" at 38,239 size 120x40; TextOff 'Tetracycline'
      on Click: ActivateScreen("4_ORDER", 0); SetTag("Selected_URL", 'file:///C:/ASRS_Video/clip261.html')
      on Activate: SetTag("Selected_Medicine", 261)
      on Release: SetTag("ยา 261", 0)
      on Press: SetTag("ยา 261", 1)
   Button "Button_9" at 688,16 size 96x40; TextOff 'Next'
      on Press: ActivateScreen("6_1", 0)
   Button "Button_10" at 38,415 size 120x40; TextOff 'Norfloxacin'
      on Click: ActivateScreen("4_ORDER", 0); SetTag("Selected_URL", 'file:///C:/ASRS_Video/clip266.html')
      on Activate: SetTag("Selected_Medicine", 266)
      on Release: SetTag("ยา 266", 0)
      on Press: SetTag("ยา 266", 1)
   Button "Button_2" at 189,240 size 120x40; TextOff 'Minocycline'
      on Click: ActivateScreen("4_ORDER", 0); SetTag("Selected_URL", 'file:///C:/ASRS_Video/clip262.html')
      on Activate: SetTag("Selected_Medicine", 262)
      on Release: SetTag("ยา 262", 0)
      on Press: SetTag("ยา 262", 1)
   Button "Button_3" at 190,415 size 120x40; TextOff 'Ofloxacin'
      on Click: ActivateScreen("4_ORDER", 0); SetTag("Selected_URL", 'file:///C:/ASRS_Video/clip267.html')
      on Activate: SetTag("Selected_Medicine", 267)
      on Release: SetTag("ยา 267", 0)
      on Press: SetTag("ยา 267", 1)
   Button "Button_4" at 340,240 size 120x40; TextOff 'Ciprofloxacin'
      on Click: ActivateScreen("4_ORDER", 0); SetTag("Selected_URL", 'file:///C:/ASRS_Video/clip263.html')
      on Activate: SetTag("Selected_Medicine", 263)
      on Release: SetTag("ยา 263", 0)
      on Press: SetTag("ยา 263", 1)
   Button "Button_5" at 340,416 size 120x40; TextOff 'Co-trimoxazole'
      on Click: ActivateScreen("4_ORDER", 0); SetTag("Selected_URL", 'file:///C:/ASRS_Video/clip268.html')
      on Activate: SetTag("Selected_Medicine", 268)
      on Release: SetTag("ยา 268", 0)
      on Press: SetTag("ยา 268", 1)
   Button "Button_6" at 492,416 size 120x40; TextOff 'Sulfadiazine'
      on Click: ActivateScreen("4_ORDER", 0); SetTag("Selected_URL", 'file:///C:/ASRS_Video/clip269.html')
      on Activate: SetTag("Selected_Medicine", 269)
      on Release: SetTag("ยา 269", 0)
      on Press: SetTag("ยา 269", 1)
   Button "Button_7" at 492,240 size 120x40; TextOff 'Levofloxacin'
      on Click: ActivateScreen("4_ORDER", 0); SetTag("Selected_URL", 'file:///C:/ASRS_Video/clip264.html')
      on Activate: SetTag("Selected_Medicine", 264)
      on Release: SetTag("ยา 264", 0)
      on Press: SetTag("ยา 264", 1)
   Button "Button_8" at 644,240 size 120x40; TextOff 'Moxifloxacin'
      on Click: ActivateScreen("4_ORDER", 0); SetTag("Selected_URL", 'file:///C:/ASRS_Video/clip265.html')
      on Activate: SetTag("Selected_Medicine", 265)
      on Release: SetTag("ยา 265", 0)
      on Press: SetTag("ยา 265", 1)
   Button "Button_11" at 645,416 size 120x40; TextOff 'Sulfasalazine'
      on Click: ActivateScreen("4_ORDER", 0); SetTag("Selected_URL", 'file:///C:/ASRS_Video/clip270.html')
      on Activate: SetTag("Selected_Medicine", 270)
      on Release: SetTag("ยา 270", 0)
      on Press: SetTag("ยา 270", 1)
   Button "Button_12" at 24,16 size 94x40; TextOff 'Back'
      on Press: ActivateScreen("4_1", 0)
   GraphicView "Template_Graphic view_1" at 693,20 size 36x32; Picture "play"
   GraphicView "Template_Graphic view_2" at 27,19 size 36x32; Picture "fast-backward"
   GraphicView "Template_Graphic view_3" at 37,128 size 120x104; Picture "41"
   GraphicView "Template_Graphic view_4" at 191,129 size 120x104; Picture "42"
   GraphicView "Template_Graphic view_5" at 339,129 size 120x104; Picture "43"
   GraphicView "Template_Graphic view_6" at 493,129 size 120x104; Picture "44"
   GraphicView "Template_Graphic view_7" at 645,129 size 120x104; Picture "45"
   GraphicView "Template_Graphic view_8" at 38,305 size 120x104; Picture "46"
   GraphicView "Template_Graphic view_9" at 189,304 size 120x112; Picture "47"
   GraphicView "Template_Graphic view_10" at 351,307 size 96x104; Picture "48"
   GraphicView "Template_Graphic view_11" at 497,304 size 120x112; Picture "49"
   GraphicView "Template_Graphic view_12" at 645,304 size 120x104; Picture "50"
   TextField "Template_Text field_2" at 201,80 size 20x32; Text '5'

screen "6_1" 800x480, template "Template_2"
   Button "Button_1" at 38,239 size 120x40; TextOff 'Metronidazole'
      on Click: ActivateScreen("4_ORDER", 0); SetTag("Selected_URL", 'file:///C:/ASRS_Video/clip271.html')
      on Activate: SetTag("Selected_Medicine", 271)
      on Release: SetTag("ยา 271", 0)
      on Press: SetTag("ยา 271", 1)
   Button "Button_9" at 688,16 size 96x40; TextOff 'Next'
      on Press: ActivateScreen("7_1", 0)
   Button "Button_10" at 38,415 size 120x40; TextOff 'Isoniazid'
      on Click: ActivateScreen("4_ORDER", 0); SetTag("Selected_URL", 'file:///C:/ASRS_Video/clip276.html')
      on Activate: SetTag("Selected_Medicine", 276)
      on Release: SetTag("ยา 276", 0)
      on Press: SetTag("ยา 276", 1)
   Button "Button_2" at 189,240 size 120x40; TextOff 'Tinidazole'
      on Click: ActivateScreen("4_ORDER", 0); SetTag("Selected_URL", 'file:///C:/ASRS_Video/clip272.html')
      on Activate: SetTag("Selected_Medicine", 272)
      on Release: SetTag("ยา 272", 0)
      on Press: SetTag("ยา 272", 1)
   Button "Button_3" at 190,415 size 120x40; TextOff 'Ethambutol'
      on Click: ActivateScreen("4_ORDER", 0); SetTag("Selected_URL", 'file:///C:/ASRS_Video/clip277.html')
      on Activate: SetTag("Selected_Medicine", 277)
      on Release: SetTag("ยา 277", 0)
      on Press: SetTag("ยา 277", 1)
   Button "Button_4" at 340,240 size 120x40; TextOff 'Nitrofurantoin'
      on Click: ActivateScreen("4_ORDER", 0); SetTag("Selected_URL", 'file:///C:/ASRS_Video/clip273.html')
      on Activate: SetTag("Selected_Medicine", 273)
      on Release: SetTag("ยา 273", 0)
      on Press: SetTag("ยา 273", 1)
   Button "Button_5" at 340,416 size 120x40; TextOff 'Pyrazinamide'
      on Click: ActivateScreen("4_ORDER", 0); SetTag("Selected_URL", 'file:///C:/ASRS_Video/clip278.html')
      on Activate: SetTag("Selected_Medicine", 288)
      on Release: SetTag("ยา 278", 0)
      on Press: SetTag("ยา 278", 1)
   Button "Button_6" at 492,416 size 120x40; TextOff 'Ethionamide'
      on Click: ActivateScreen("4_ORDER", 0); SetTag("Selected_URL", 'file:///C:/ASRS_Video/clip279.html')
      on Activate: SetTag("Selected_Medicine", 279)
      on Release: SetTag("ยา 279", 0)
      on Press: SetTag("ยา 279", 1)
   Button "Button_7" at 492,240 size 120x40; TextOff 'Fosfomycin'
      on Click: ActivateScreen("4_ORDER", 0); SetTag("Selected_URL", 'file:///C:/ASRS_Video/clip274.html')
      on Activate: SetTag("Selected_Medicine", 274)
      on Release: SetTag("ยา 274", 0)
      on Press: SetTag("ยา 274", 1)
   Button "Button_8" at 644,240 size 120x40; TextOff 'Rifampicin'
      on Click: ActivateScreen("4_ORDER", 0); SetTag("Selected_URL", 'file:///C:/ASRS_Video/clip275.html')
      on Activate: SetTag("Selected_Medicine", 275)
      on Release: SetTag("ยา 275", 0)
      on Press: SetTag("ยา 275", 1)
   Button "Button_11" at 645,416 size 120x40; TextOff 'Cycloserine'
      on Click: ActivateScreen("4_ORDER", 0); SetTag("Selected_URL", 'file:///C:/ASRS_Video/clip280.html')
      on Activate: SetTag("Selected_Medicine", 280)
      on Release: SetTag("ยา 280", 0)
      on Press: SetTag("ยา 280", 1)
   Button "Button_12" at 24,16 size 94x40; TextOff 'Back'
      on Press: ActivateScreen("5_1", 0)
   GraphicView "Template_Graphic view_1" at 693,20 size 36x32; Picture "play"
   GraphicView "Template_Graphic view_2" at 27,19 size 36x32; Picture "fast-backward"
   GraphicView "Template_Graphic view_3" at 37,128 size 120x104; Picture "51"
   GraphicView "Template_Graphic view_4" at 191,129 size 120x104; Picture "52"
   GraphicView "Template_Graphic view_5" at 339,129 size 120x104; Picture "53"
   GraphicView "Template_Graphic view_6" at 493,129 size 120x104; Picture "54"
   GraphicView "Template_Graphic view_7" at 645,129 size 120x104; Picture "55"
   GraphicView "Template_Graphic view_8" at 38,305 size 120x104; Picture "56"
   GraphicView "Template_Graphic view_9" at 189,304 size 120x112; Picture "57"
   GraphicView "Template_Graphic view_10" at 351,307 size 96x104; Picture "58"
   GraphicView "Template_Graphic view_11" at 497,304 size 120x112; Picture "59"
   GraphicView "Template_Graphic view_12" at 645,304 size 120x104; Picture "60"
   TextField "Template_Text field_2" at 201,80 size 20x32; Text '6'

screen "7_1" 800x480, template "Template_2"
   Button "Button_1" at 38,239 size 120x40; TextOff 'Fluconazole'
      on Click: ActivateScreen("4_ORDER", 0); SetTag("Selected_URL", 'file:///C:/ASRS_Video/clip281.html')
      on Activate: SetTag("Selected_Medicine", 281)
      on Release: SetTag("ยา 281", 0)
      on Press: SetTag("ยา 281", 1)
   Button "Button_9" at 688,16 size 96x40; TextOff 'Next'
      on Press: ActivateScreen("8_1", 0)
   Button "Button_10" at 38,415 size 120x40; TextOff 'Nystatin'
      on Click: ActivateScreen("4_ORDER", 0); SetTag("Selected_URL", 'file:///C:/ASRS_Video/clip286.html')
      on Activate: SetTag("Selected_Medicine", 286)
      on Release: SetTag("ยา 286", 0)
      on Press: SetTag("ยา 286", 1)
   Button "Button_2" at 189,240 size 120x40; TextOff 'Itraconazole'
      on Click: ActivateScreen("4_ORDER", 0); SetTag("Selected_URL", 'file:///C:/ASRS_Video/clip282.html')
      on Activate: SetTag("Selected_Medicine", 282)
      on Release: SetTag("ยา 282", 0)
      on Press: SetTag("ยา 282", 1)
   Button "Button_3" at 190,415 size 120x40; TextOff 'Clotrimazole'
      on Click: ActivateScreen("4_ORDER", 0); SetTag("Selected_URL", 'file:///C:/ASRS_Video/clip287.html')
      on Activate: SetTag("Selected_Medicine", 287)
      on Release: SetTag("ยา 287", 0)
      on Press: SetTag("ยา 287", 1)
   Button "Button_4" at 340,240 size 120x40; TextOff 'Ketoconazole'
      on Click: ActivateScreen("4_ORDER", 0); SetTag("Selected_URL", 'file:///C:/ASRS_Video/clip283.html')
      on Activate: SetTag("Selected_Medicine", 283)
      on Release: SetTag("ยา 283", 0)
      on Press: SetTag("ยา 283", 1)
   Button "Button_5" at 340,416 size 120x40; TextOff 'Miconazole'
      on Click: ActivateScreen("4_ORDER", 0); SetTag("Selected_URL", 'file:///C:/ASRS_Video/clip288.html')
      on Activate: SetTag("Selected_Medicine", 288)
      on Release: SetTag("ยา 288", 0)
      on Press: SetTag("ยา 288", 1)
   Button "Button_6" at 492,416 size 120x40; TextOff 'Terbinafine'
      on Click: ActivateScreen("4_ORDER", 0); SetTag("Selected_URL", 'file:///C:/ASRS_Video/clip289.html')
      on Activate: SetTag("Selected_Medicine", 289)
      on Release: SetTag("ยา 289", 0)
      on Press: SetTag("ยา 289", 1)
   Button "Button_7" at 492,240 size 120x40; TextOff 'Voriconazole'
      on Click: ActivateScreen("4_ORDER", 0); SetTag("Selected_URL", 'file:///C:/ASRS_Video/clip284.html')
      on Activate: SetTag("Selected_Medicine", 284)
      on Release: SetTag("ยา 284", 0)
      on Press: SetTag("ยา 284", 1)
   Button "Button_8" at 644,240 size 120x40; TextOff 'Amphotericin B'
      on Click: ActivateScreen("4_ORDER", 0); SetTag("Selected_URL", 'file:///C:/ASRS_Video/clip285.html')
      on Activate: SetTag("Selected_Medicine", 285)
      on Release: SetTag("ยา 285", 0)
      on Press: SetTag("ยา 285", 1)
   Button "Button_11" at 645,416 size 120x40; TextOff 'Griseofulvin'
      on Click: ActivateScreen("4_ORDER", 0); SetTag("Selected_URL", 'file:///C:/ASRS_Video/clip290.html')
      on Activate: SetTag("Selected_Medicine", 290)
      on Release: SetTag("ยา 290", 0)
      on Press: SetTag("ยา 290", 1)
   Button "Button_12" at 24,16 size 94x40; TextOff 'Back'
      on Press: ActivateScreen("6_1", 0)
   GraphicView "Template_Graphic view_1" at 693,20 size 36x32; Picture "play"
   GraphicView "Template_Graphic view_2" at 27,19 size 36x32; Picture "fast-backward"
   GraphicView "Template_Graphic view_3" at 37,128 size 120x104; Picture "61"
   GraphicView "Template_Graphic view_4" at 191,129 size 120x104; Picture "62"
   GraphicView "Template_Graphic view_5" at 339,129 size 120x104; Picture "63"
   GraphicView "Template_Graphic view_6" at 493,129 size 120x104; Picture "64"
   GraphicView "Template_Graphic view_7" at 645,129 size 120x104; Picture "65"
   GraphicView "Template_Graphic view_8" at 38,305 size 120x104; Picture "66"
   GraphicView "Template_Graphic view_9" at 189,304 size 120x104; Picture "67"
   GraphicView "Template_Graphic view_10" at 351,307 size 96x104; Picture "68"
   GraphicView "Template_Graphic view_11" at 497,304 size 120x112; Picture "69"
   GraphicView "Template_Graphic view_12" at 645,304 size 120x104; Picture "70"
   TextField "Template_Text field_2" at 201,80 size 20x32; Text '7'
   TextField "Text field_1" at 0,0 size 101x22; Text 'Amphotericin B'

